Staubli VAL3: io.pjx

--- io.pjx ---
Parameters version=s8.10.3Cs9_BS2093 stackSize=5000 millimeterUnit=true
Program file=commentIO.pgx
Program file=getAnaIO.pgx
Program file=getAngIOSize.pgx
Program file=getDigIO.pgx
Program file=getDigIOSize.pgx
Program file=init.pgx
Program file=linkIO.pgx
Program file=linkStatusIO.pgx
Program file=resetBusSelect.pgx
Program file=setAnaOutput.pgx
Program file=setAngINList.pgx
Program file=setAngOUTList.pgx
Program file=setDigOutNoAlm.pgx
Program file=setDigOutput.pgx
Program file=start.pgx
Program file=stop.pgx
Program file=waitAnaInput.pgx
Program file=waitDigInput.pgx
Data file=io.dtx
Library alias=rs path=Disk://source/projectSource/robotStatus/robotStatus.pjx
Type name=dioItem path=Disk://source/template/dioItem/dioItem.pjx
Type name=aioItem path=Disk://source/template/aioItem/aioItem.pjx

--- io.dtx ---
public aio _aInEthercat[16]
public aio _aInEthernet[20]
public aio _aInModbus[16]
public aio _aInProfibus[16]
public aio _aInProfinet[8]
  [0] = {link=61F414E4-CB2A-4A4A-A70F-3C6D612AB3AA}
  [1] = {link=443D484E-60E0-45BD-99C4-97873755DFDA}
  [2] = {link=73C25A3F-C0C4-4812-B693-CDA309C2D933}
  [3] = {link=D3F549A9-B3EA-403D-BF4C-7070E9F5D37B}
  [4] = {link=F3F4C9C0-1F7C-4DDD-AA59-2014D98A0E36}
  [5] = {link=64B8C6E8-3A71-49B0-BD71-5728B0329AAB}
  [6] = {link=218C656F-9E2A-4E1B-B485-E83EC4F0FE99}
  [7] = {link=66AABE0A-89B4-481F-83AB-C514130625BA}
public aio _aInUser[16]
public aio _aOEthercat[16]
public aio _aOEthernet[20]
public aio _aOModbus[16]
public aio _aOProfibus[16]
public aio _aOProfinet[8]
  [0] = {link=5FFE21EC-528D-4C47-A8D5-7C4CFC474629}
  [1] = {link=6C0C10F5-5D52-4306-AECC-A9DCF4E15FA5}
  [2] = {link=96FBB4C4-7B28-4C73-AFB9-CDBD1E0FA505}
  [3] = {link=3CD60215-4462-490B-9BA1-05C4B27AD9CF}
  [4] = {link=45C44C09-08B8-4891-969D-45390D63770F}
  [5] = {link=DD02F8D1-5F5E-4FDF-BD15-7DB79F0068FE}
  [6] = {link=0578226E-4341-48AC-B576-D095F8D3C1C5}
  [7] = {link=D8473422-71DA-4369-901E-04429E7E73E1}
public aio _aOutUser[16]
public aio aInJobNumber
public aio aInVirtual[24]
  [0] = {link=VirtualIOBoards\VirtualBoard0\%IF128}
  [1] = {link=VirtualIOBoards\VirtualBoard0\%IF160}
  [2] = {link=VirtualIOBoards\VirtualBoard0\%IF192}
  [3] = {link=VirtualIOBoards\VirtualBoard0\%IF224}
  [4] = {link=VirtualIOBoards\VirtualBoard0\%IF256}
  [5] = {link=VirtualIOBoards\VirtualBoard0\%IF288}
  [6] = {link=VirtualIOBoards\VirtualBoard0\%IF320}
  [7] = {link=VirtualIOBoards\VirtualBoard0\%IF352}
  [8] = {link=VirtualIOBoards\VirtualBoard0\%IF384}
  [9] = {link=VirtualIOBoards\VirtualBoard0\%IF416}
  [10] = {link=VirtualIOBoards\VirtualBoard0\%IF448}
  [11] = {link=VirtualIOBoards\VirtualBoard0\%IF480}
  [12] = {link=VirtualIOBoards\VirtualBoard0\%IF512}
  [13] = {link=VirtualIOBoards\VirtualBoard0\%IF544}
  [14] = {link=VirtualIOBoards\VirtualBoard0\%IF576}
  [15] = {link=VirtualIOBoards\VirtualBoard0\%IF608}
  [16] = {link=VirtualIOBoards\VirtualBoard0\%IF640}
  [17] = {link=VirtualIOBoards\VirtualBoard0\%IF672}
  [18] = {link=VirtualIOBoards\VirtualBoard0\%IF704}
  [19] = {link=VirtualIOBoards\VirtualBoard0\%IF736}
  [20] = {link=VirtualIOBoards\VirtualBoard0\%IF768}
  [21] = {link=VirtualIOBoards\VirtualBoard0\%IF800}
  [22] = {link=VirtualIOBoards\VirtualBoard0\%IF832}
  [23] = {link=VirtualIOBoards\VirtualBoard0\%IF864}
public aio aInput[8]
  [0] = {link=61F414E4-CB2A-4A4A-A70F-3C6D612AB3AA}
  [1] = {link=443D484E-60E0-45BD-99C4-97873755DFDA}
  [2] = {link=73C25A3F-C0C4-4812-B693-CDA309C2D933}
  [3] = {link=D3F549A9-B3EA-403D-BF4C-7070E9F5D37B}
  [4] = {link=F3F4C9C0-1F7C-4DDD-AA59-2014D98A0E36}
  [5] = {link=64B8C6E8-3A71-49B0-BD71-5728B0329AAB}
  [6] = {link=218C656F-9E2A-4E1B-B485-E83EC4F0FE99}
  [7] = {link=66AABE0A-89B4-481F-83AB-C514130625BA}
public aio aOutJobNumber
public aio aOutVirtual[24]
  [0] = {link=VirtualIOBoards\VirtualBoard0\%QF128}
  [1] = {link=VirtualIOBoards\VirtualBoard0\%QF160}
  [2] = {link=VirtualIOBoards\VirtualBoard0\%QF192}
  [3] = {link=VirtualIOBoards\VirtualBoard0\%QF224}
  [4] = {link=VirtualIOBoards\VirtualBoard0\%QF256}
  [5] = {link=VirtualIOBoards\VirtualBoard0\%QF288}
  [6] = {link=VirtualIOBoards\VirtualBoard0\%QF320}
  [7] = {link=VirtualIOBoards\VirtualBoard0\%QF352}
  [8] = {link=VirtualIOBoards\VirtualBoard0\%QF384}
  [9] = {link=VirtualIOBoards\VirtualBoard0\%QF416}
  [10] = {link=VirtualIOBoards\VirtualBoard0\%QF448}
  [11] = {link=VirtualIOBoards\VirtualBoard0\%QF480}
  [12] = {link=VirtualIOBoards\VirtualBoard0\%QF512}
  [13] = {link=VirtualIOBoards\VirtualBoard0\%QF544}
  [14] = {link=VirtualIOBoards\VirtualBoard0\%QF576}
  [15] = {link=VirtualIOBoards\VirtualBoard0\%QF608}
  [16] = {link=VirtualIOBoards\VirtualBoard0\%QF640}
  [17] = {link=VirtualIOBoards\VirtualBoard0\%QF672}
  [18] = {link=VirtualIOBoards\VirtualBoard0\%QF704}
  [19] = {link=VirtualIOBoards\VirtualBoard0\%QF736}
  [20] = {link=VirtualIOBoards\VirtualBoard0\%QF768}
  [21] = {link=VirtualIOBoards\VirtualBoard0\%QF800}
  [22] = {link=VirtualIOBoards\VirtualBoard0\%QF832}
  [23] = {link=VirtualIOBoards\VirtualBoard0\%QF864}
public aio aOutput[8]
  [0] = {link=5FFE21EC-528D-4C47-A8D5-7C4CFC474629}
  [1] = {link=6C0C10F5-5D52-4306-AECC-A9DCF4E15FA5}
  [2] = {link=96FBB4C4-7B28-4C73-AFB9-CDBD1E0FA505}
  [3] = {link=3CD60215-4462-490B-9BA1-05C4B27AD9CF}
  [4] = {link=45C44C09-08B8-4891-969D-45390D63770F}
  [5] = {link=DD02F8D1-5F5E-4FDF-BD15-7DB79F0068FE}
  [6] = {link=0578226E-4341-48AC-B576-D095F8D3C1C5}
  [7] = {link=D8473422-71DA-4369-901E-04429E7E73E1}
public aioItem aInItem[8]
  [0]
    aio aAio = {link=61F414E4-CB2A-4A4A-A70F-3C6D612AB3AA}
    string sComment = "接收程序号"
  [1]
    aio aAio = {link=443D484E-60E0-45BD-99C4-97873755DFDA}
    string sComment = "刷子号反馈"
  [2]
    aio aAio = {link=73C25A3F-C0C4-4812-B693-CDA309C2D933}
    string sComment = "备用"
  [3]
    aio aAio = {link=D3F549A9-B3EA-403D-BF4C-7070E9F5D37B}
    string sComment = "备用"
  [4]
    aio aAio = {link=F3F4C9C0-1F7C-4DDD-AA59-2014D98A0E36}
    string sComment = "备用"
  [5]
    aio aAio = {link=64B8C6E8-3A71-49B0-BD71-5728B0329AAB}
    string sComment = "备用"
  [6]
    aio aAio = {link=218C656F-9E2A-4E1B-B485-E83EC4F0FE99}
    string sComment = "备用"
  [7]
    aio aAio = {link=66AABE0A-89B4-481F-83AB-C514130625BA}
    string sComment = "备用"
public aioItem aOutItem[8]
  [0]
    aio aAio = {link=5FFE21EC-528D-4C47-A8D5-7C4CFC474629}
    string sComment = "程序号反馈"
  [1]
    aio aAio = {link=6C0C10F5-5D52-4306-AECC-A9DCF4E15FA5}
    string sComment = "刷子号"
  [2]
    aio aAio = {link=96FBB4C4-7B28-4C73-AFB9-CDBD1E0FA505}
    string sComment = "备用"
  [3]
    aio aAio = {link=3CD60215-4462-490B-9BA1-05C4B27AD9CF}
    string sComment = "备用"
  [4]
    aio aAio = {link=45C44C09-08B8-4891-969D-45390D63770F}
    string sComment = "备用"
  [5]
    aio aAio = {link=DD02F8D1-5F5E-4FDF-BD15-7DB79F0068FE}
    string sComment = "备用"
  [6]
    aio aAio = {link=0578226E-4341-48AC-B576-D095F8D3C1C5}
    string sComment = "备用"
  [7]
    aio aAio = {link=D8473422-71DA-4369-901E-04429E7E73E1}
    string sComment = "备用"
bool bBusSelect[6]
bool bUseAnalog = true
public dio _dInEtherCat[96]
public dio _dInEtherNet[128]
  [0] = {link=3C99ACBA-F1D4-4A68-A21C-89A8C66262F3}
  [1] = {link=A8C10724-75A9-4217-88F5-3321E2E2ACAD}
  [2] = {link=3FECD266-02DB-40D3-AA00-852A922114D7}
  [3] = {link=527ABC03-504A-4B4E-8384-0B648B30A7EE}
  [4] = {link=F6BC421B-A283-4F49-B66E-4A61065D35DB}
  [5] = {link=AF78B140-D810-4E0E-A464-37CD3BF21C1F}
  [6] = {link=54025B48-0E34-4C00-83F4-7C1C00C78D0E}
  [7] = {link=C893EABF-80A0-4CC4-8CB1-35D77AC88EDF}
  [8] = {link=B91BA001-E4EA-48BD-931D-F38D504579C9}
  [9] = {link=F2BD5778-F2D0-400E-8EB0-EB74F7A1D168}
  [10] = {link=00F50513-209B-4FEC-BCA0-2732338E58E1}
  [11] = {link=881EE622-97CE-4B32-A64C-C6F69EF3ED05}
  [12] = {link=56AD774C-0018-466F-B601-292CE44541BC}
  [13] = {link=4324DB33-706B-4D11-8D24-EAF877265392}
  [14] = {link=5AF359B1-8E78-40AA-A03B-F8A0077C8703}
  [15] = {link=ApplicomIO-1\PFN-IN\%I0[15]}
  [16] = {link=ApplicomIO-1\PFN-IN\%I0[16]}
  [17] = {link=ApplicomIO-1\PFN-IN\%I0[17]}
  [18] = {link=ApplicomIO-1\PFN-IN\%I0[18]}
  [19] = {link=ApplicomIO-1\PFN-IN\%I0[19]}
  [20] = {link=ApplicomIO-1\PFN-IN\%I0[20]}
  [21] = {link=ApplicomIO-1\PFN-IN\%I0[21]}
  [22] = {link=ApplicomIO-1\PFN-IN\%I0[22]}
  [23] = {link=ApplicomIO-1\PFN-IN\%I0[23]}
  [24] = {link=ApplicomIO-1\PFN-IN\%I0[24]}
  [25] = {link=ApplicomIO-1\PFN-IN\%I0[25]}
  [26] = {link=ApplicomIO-1\PFN-IN\%I0[26]}
  [27] = {link=ApplicomIO-1\PFN-IN\%I0[27]}
  [28] = {link=ApplicomIO-1\PFN-IN\%I0[28]}
  [29] = {link=ApplicomIO-1\PFN-IN\%I0[29]}
  [30] = {link=ApplicomIO-1\PFN-IN\%I0[30]}
  [31] = {link=ApplicomIO-1\PFN-IN\%I0[31]}
  [32] = {link=ApplicomIO-1\PFN-IN\%I0[32]}
  [33] = {link=ApplicomIO-1\PFN-IN\%I0[33]}
  [34] = {link=ApplicomIO-1\PFN-IN\%I0[34]}
  [35] = {link=ApplicomIO-1\PFN-IN\%I0[35]}
  [36] = {link=ApplicomIO-1\PFN-IN\%I0[36]}
  [37] = {link=ApplicomIO-1\PFN-IN\%I0[37]}
  [38] = {link=ApplicomIO-1\PFN-IN\%I0[38]}
  [39] = {link=ApplicomIO-1\PFN-IN\%I0[39]}
  [40] = {link=ApplicomIO-1\PFN-IN\%I0[40]}
  [41] = {link=ApplicomIO-1\PFN-IN\%I0[41]}
  [42] = {link=ApplicomIO-1\PFN-IN\%I0[42]}
  [43] = {link=ApplicomIO-1\PFN-IN\%I0[43]}
  [44] = {link=ApplicomIO-1\PFN-IN\%I0[44]}
  [45] = {link=ApplicomIO-1\PFN-IN\%I0[45]}
  [46] = {link=ApplicomIO-1\PFN-IN\%I0[46]}
  [47] = {link=ApplicomIO-1\PFN-IN\%I0[47]}
  [48] = {link=ApplicomIO-1\PFN-IN\%I0[48]}
  [49] = {link=ApplicomIO-1\PFN-IN\%I0[49]}
  [50] = {link=ApplicomIO-1\PFN-IN\%I0[50]}
  [51] = {link=ApplicomIO-1\PFN-IN\%I0[51]}
  [52] = {link=ApplicomIO-1\PFN-IN\%I0[52]}
  [53] = {link=ApplicomIO-1\PFN-IN\%I0[53]}
  [54] = {link=ApplicomIO-1\PFN-IN\%I0[54]}
  [55] = {link=ApplicomIO-1\PFN-IN\%I0[55]}
  [56] = {link=ApplicomIO-1\PFN-IN\%I0[56]}
  [57] = {link=ApplicomIO-1\PFN-IN\%I0[57]}
  [58] = {link=ApplicomIO-1\PFN-IN\%I0[58]}
  [59] = {link=ApplicomIO-1\PFN-IN\%I0[59]}
  [60] = {link=ApplicomIO-1\PFN-IN\%I0[60]}
  [61] = {link=ApplicomIO-1\PFN-IN\%I0[61]}
  [62] = {link=ApplicomIO-1\PFN-IN\%I0[62]}
  [63] = {link=ApplicomIO-1\PFN-IN\%I0[63]}
public dio _dInModbus[96]
public dio _dInProfibus[96]
  [0] = {link=ApplicomIO-1\PFB-BLOCK\%I0[0]}
  [1] = {link=ApplicomIO-1\PFB-BLOCK\%I0[1]}
  [2] = {link=ApplicomIO-1\PFB-BLOCK\%I0[2]}
  [3] = {link=ApplicomIO-1\PFB-BLOCK\%I0[3]}
  [4] = {link=ApplicomIO-1\PFB-BLOCK\%I0[4]}
  [5] = {link=ApplicomIO-1\PFB-BLOCK\%I0[5]}
  [6] = {link=ApplicomIO-1\PFB-BLOCK\%I0[6]}
  [7] = {link=ApplicomIO-1\PFB-BLOCK\%I0[7]}
  [8] = {link=ApplicomIO-1\PFB-BLOCK\%I0[8]}
  [9] = {link=ApplicomIO-1\PFB-BLOCK\%I0[9]}
  [10] = {link=ApplicomIO-1\PFB-BLOCK\%I0[10]}
  [11] = {link=ApplicomIO-1\PFB-BLOCK\%I0[11]}
  [12] = {link=ApplicomIO-1\PFB-BLOCK\%I0[12]}
  [13] = {link=ApplicomIO-1\PFB-BLOCK\%I0[13]}
  [14] = {link=ApplicomIO-1\PFB-BLOCK\%I0[14]}
  [15] = {link=ApplicomIO-1\PFB-BLOCK\%I0[15]}
  [16] = {link=ApplicomIO-1\PFB-BLOCK\%I0[16]}
  [17] = {link=ApplicomIO-1\PFB-BLOCK\%I0[17]}
  [18] = {link=ApplicomIO-1\PFB-BLOCK\%I0[18]}
  [19] = {link=ApplicomIO-1\PFB-BLOCK\%I0[19]}
  [20] = {link=ApplicomIO-1\PFB-BLOCK\%I0[20]}
  [21] = {link=ApplicomIO-1\PFB-BLOCK\%I0[21]}
  [22] = {link=ApplicomIO-1\PFB-BLOCK\%I0[22]}
  [23] = {link=ApplicomIO-1\PFB-BLOCK\%I0[23]}
  [24] = {link=ApplicomIO-1\PFB-BLOCK\%I0[24]}
  [25] = {link=ApplicomIO-1\PFB-BLOCK\%I0[25]}
  [26] = {link=ApplicomIO-1\PFB-BLOCK\%I0[26]}
  [27] = {link=ApplicomIO-1\PFB-BLOCK\%I0[27]}
  [28] = {link=ApplicomIO-1\PFB-BLOCK\%I0[28]}
  [29] = {link=ApplicomIO-1\PFB-BLOCK\%I0[29]}
  [30] = {link=ApplicomIO-1\PFB-BLOCK\%I0[30]}
  [31] = {link=ApplicomIO-1\PFB-BLOCK\%I0[31]}
  [32] = {link=ApplicomIO-1\PFB-BLOCK\%I0[32]}
  [33] = {link=ApplicomIO-1\PFB-BLOCK\%I0[33]}
  [34] = {link=ApplicomIO-1\PFB-BLOCK\%I0[34]}
  [35] = {link=ApplicomIO-1\PFB-BLOCK\%I0[35]}
  [36] = {link=ApplicomIO-1\PFB-BLOCK\%I0[36]}
  [37] = {link=ApplicomIO-1\PFB-BLOCK\%I0[37]}
  [38] = {link=ApplicomIO-1\PFB-BLOCK\%I0[38]}
  [39] = {link=ApplicomIO-1\PFB-BLOCK\%I0[39]}
  [40] = {link=ApplicomIO-1\PFB-BLOCK\%I0[40]}
  [41] = {link=ApplicomIO-1\PFB-BLOCK\%I0[41]}
  [42] = {link=ApplicomIO-1\PFB-BLOCK\%I0[42]}
  [43] = {link=ApplicomIO-1\PFB-BLOCK\%I0[43]}
  [44] = {link=ApplicomIO-1\PFB-BLOCK\%I0[44]}
  [45] = {link=ApplicomIO-1\PFB-BLOCK\%I0[45]}
  [46] = {link=ApplicomIO-1\PFB-BLOCK\%I0[46]}
  [47] = {link=ApplicomIO-1\PFB-BLOCK\%I0[47]}
  [48] = {link=ApplicomIO-1\PFB-BLOCK\%I0[48]}
  [49] = {link=ApplicomIO-1\PFB-BLOCK\%I0[49]}
  [50] = {link=ApplicomIO-1\PFB-BLOCK\%I0[50]}
  [51] = {link=ApplicomIO-1\PFB-BLOCK\%I0[51]}
  [52] = {link=ApplicomIO-1\PFB-BLOCK\%I0[52]}
  [53] = {link=ApplicomIO-1\PFB-BLOCK\%I0[53]}
  [54] = {link=ApplicomIO-1\PFB-BLOCK\%I0[54]}
  [55] = {link=ApplicomIO-1\PFB-BLOCK\%I0[55]}
  [56] = {link=ApplicomIO-1\PFB-BLOCK\%I0[56]}
  [57] = {link=ApplicomIO-1\PFB-BLOCK\%I0[57]}
  [58] = {link=ApplicomIO-1\PFB-BLOCK\%I0[58]}
  [59] = {link=ApplicomIO-1\PFB-BLOCK\%I0[59]}
  [60] = {link=ApplicomIO-1\PFB-BLOCK\%I0[60]}
  [61] = {link=ApplicomIO-1\PFB-BLOCK\%I0[61]}
  [62] = {link=ApplicomIO-1\PFB-BLOCK\%I0[62]}
  [63] = {link=ApplicomIO-1\PFB-BLOCK\%I0[63]}
public dio _dInProfinet[128]
  [0] = {link=801699AD-0D4E-40AF-A7AF-E7C40311637E}
  [1] = {link=842E3CE8-5982-430F-AA8E-B2F701DC178B}
  [2] = {link=F299EF97-EDDD-4BB8-AA07-719E60051D06}
  [3] = {link=0D6C59A5-572E-4845-9D24-D0618D782DD4}
  [4] = {link=CC171C2B-47CE-4C45-9659-7FCDC013CE94}
  [5] = {link=1A1317E2-9651-45BA-ACEA-D1820BFA9703}
  [6] = {link=1B720B0E-A94A-4B35-8241-512C8CFE7420}
  [7] = {link=6F68113A-0DD2-4F74-B0DE-02F63C641B3D}
  [8] = {link=DB25555B-9639-404C-BF41-A1E4182E7853}
  [9] = {link=A68ADCD7-077C-45ED-AE36-CA1771248567}
  [10] = {link=3971923C-046E-4FB8-8CDF-8298982DD00B}
  [11] = {link=C253DB67-AB15-493D-BA5F-F7404DA89E40}
  [12] = {link=5F58F424-9E7E-46E6-B5AD-37E850D30CCF}
  [13] = {link=0B266260-B4AD-4902-9CA8-DAC05E19210B}
  [14] = {link=20B44CE4-2E83-403B-A39C-4F8E5CA01265}
  [15] = {link=CD23C02B-CC02-4E28-82D0-6EB1534712A8}
  [16] = {link=550C0093-735F-4929-AB88-92E210EEA585}
  [17] = {link=58675BC9-A902-44A6-9D1E-CDCDD371E5BF}
  [18] = {link=C6C06F3F-E54C-4EE8-B5A1-0B392CB95D19}
  [19] = {link=E7996F97-FFB6-4A1D-8389-FC391F807530}
  [20] = {link=545E5659-957E-409A-983D-845A312BF10F}
  [21] = {link=896C2D61-98DD-43B3-A9FF-B63B82E13F66}
  [22] = {link=CB058ED0-A460-493F-ACD8-83515F19CB22}
  [23] = {link=8EC8BEC8-3882-4E09-82EB-ED6F4043F345}
  [24] = {link=6614FE1F-5D84-418F-8C43-3AD6E08D9885}
  [25] = {link=A0D729AE-192B-4443-98B3-A6978F97C45B}
  [26] = {link=8274EAD0-4711-40CE-9532-B3E4F6D5E848}
  [27] = {link=A4D7A453-0050-4322-BCBB-255C4251B0BA}
  [28] = {link=0CFB91EB-8B07-41BC-89A1-F8BBECCF0624}
  [29] = {link=4F7299CD-79A3-4FE2-8435-19083E83C2B9}
  [30] = {link=E49B7D09-65F8-4955-B810-3C508C434830}
  [31] = {link=2BAB1321-D2BB-48C2-8DEA-1230FF1A9D85}
  [32] = {link=C00D5C02-BF78-4EF5-B868-C5B31E42BE7F}
  [33] = {link=96859C69-E3EF-4F26-913D-E25096C13C5F}
  [34] = {link=7920EEE9-3DBF-43F3-9541-7FBE207ECE53}
  [35] = {link=1DB9160A-F63F-4C13-93B5-492FEDD177E2}
  [36] = {link=1FC4D9B1-EE44-4A9B-A22D-5889BB08EE1E}
  [37] = {link=BF970AFE-565C-4857-97A6-5A54DDAE79B6}
  [38] = {link=F909C748-B7A8-4470-A6FD-BA1A46FE4E68}
  [39] = {link=8517CD21-2BAD-4F53-9136-89235F4060C6}
  [40] = {link=6DDBB7AB-AC7B-4F3D-A091-1238925E0448}
  [41] = {link=C3CF7374-59EF-4029-99B4-FC98E25808BB}
  [42] = {link=90C02E77-8235-444D-99EB-D816EF90AFE5}
  [43] = {link=E44556E2-741A-40A0-89B2-8E32677B3EB1}
  [44] = {link=D8AFCC23-6F61-4ADD-8DE3-3FE1547AD28D}
  [45] = {link=98BC2888-38BC-4A33-A762-BDEC3E36173F}
  [46] = {link=A24DA26D-2F10-46AE-809B-0B04336865AA}
  [47] = {link=04D21FA2-EBE1-4E66-8338-7CB17174A724}
  [48] = {link=E766472B-9569-4911-A858-6F7708718D01}
  [49] = {link=92C360C1-157E-40E1-9184-03D53ECDF3F7}
  [50] = {link=6E33B145-BAC8-48E7-A184-E5A9D90B515B}
  [51] = {link=D5FDB290-CB76-4852-8AF4-F9B6FA5D3E2D}
  [52] = {link=547C3630-B2EA-42F8-AB37-EEB4C81AA149}
  [53] = {link=A60C469C-4F75-4C30-9347-66365041DE79}
  [54] = {link=6E14BCEF-8B69-4038-B259-0EF712D2AB66}
  [55] = {link=B19F0E1B-CE25-49C3-9ED7-92404708DBC9}
  [56] = {link=AFC49D6D-7F53-41F5-8159-6058E9291542}
  [57] = {link=BB08126F-937C-4C50-9A1C-252CB13BB25C}
  [58] = {link=15BF4171-EFAA-47B7-BEF9-A698BE11011C}
  [59] = {link=9A261803-1F52-41D2-8355-1C79BF1BB94D}
  [60] = {link=18F63136-91BD-4FEE-8DA3-2AA9D2E8FFA8}
  [61] = {link=55E89D2C-C808-4026-99D2-85E324C475F9}
  [62] = {link=45535323-0512-46DB-8EB0-4BF3F55D73C7}
  [63] = {link=23943399-CEE5-49D9-BFD9-55B5920F548B}
  [64] = {link=364F41EB-6BA1-4700-BD0A-C2236839044E}
  [65] = {link=96EFCAAE-6B9A-4070-B9EC-2035BA94CCB3}
  [66] = {link=FD79DB68-803F-47E7-8305-8CFFFE519C88}
  [67] = {link=82CF98E3-5511-4523-9501-B4BBAD9DC96D}
  [68] = {link=43A446B7-3C25-4DD5-9597-27365DBE2539}
  [69] = {link=01367322-9745-4163-BFB8-DF881D521F4A}
  [70] = {link=1F635259-38C5-4AB2-B093-ADA4F82FD92B}
  [71] = {link=80065B3A-E7EF-4B6D-A30A-AC2F8A1FF9BD}
  [72] = {link=138692BF-FCCE-4B34-B0E8-8C4B22C67F12}
  [73] = {link=2F598E66-6704-43A6-A433-14D902C15D10}
  [74] = {link=3D7C9642-411B-40D3-B3B9-C83D24259AF4}
  [75] = {link=2E14C0AE-1F04-4256-8959-DEAD28BB69AE}
  [76] = {link=D90512A1-D0E1-41B2-8294-59D7C1ADD8E0}
  [77] = {link=F9EFA2A2-C655-4B55-8F3F-AAE77A6FD751}
  [78] = {link=8C43F822-1313-4C63-84D2-76D62B96A58F}
  [79] = {link=0BE51982-5E8E-4776-A637-0836608FA4D4}
  [80] = {link=5CC26A0C-A759-4F9D-9C90-7643106A4280}
  [81] = {link=6B2348DB-D0C3-44B1-96EA-09FBC0D6D1F3}
  [82] = {link=091DC27E-E2EB-463E-8E4B-08B48E663650}
  [83] = {link=EC5520D5-F711-48B3-AE90-97344DDBEE5C}
  [84] = {link=E02811C8-C36E-4E92-B28C-81A727813C5B}
  [85] = {link=39EB69C5-9612-415D-9A77-D013E3B8CFD4}
  [86] = {link=FD4FFC3C-593A-4304-8BB2-18534DB95237}
  [87] = {link=D2ECCFF1-C6D1-48A4-B3A9-F333711A9798}
  [88] = {link=13EA7043-3380-41E5-9177-AAC787C21C39}
  [89] = {link=5475660F-31B7-47C3-808C-FBAB066EFE6D}
  [90] = {link=93D7CC16-1244-4B9F-85C2-564B516A38A6}
  [91] = {link=A2A5B44E-CAC8-47F1-A810-875EED5095FB}
  [92] = {link=2F9951E4-3414-412E-A45B-55B5D632DA1B}
  [93] = {link=916866A1-8E9C-42B7-A695-7CB9D795E148}
  [94] = {link=CA3200CB-BA9D-4435-B593-6CDDBB86F10C}
  [95] = {link=49AC3AF5-F49B-42A1-90B2-5DB7D6C7E051}
  [96] = {link=64E7B72A-8AE1-43E7-9A21-FF4DABD03910}
  [97] = {link=7BA0757A-43B7-4994-86FC-1740DE8C159E}
  [98] = {link=5ACF5B88-9BD6-435A-8F3F-752FE88E7935}
  [99] = {link=70DFB9C6-9CA4-44C9-8464-A31BA0D039F5}
  [100] = {link=55D5D0F9-E23A-40DA-9955-6BCB63B37099}
  [101] = {link=1AB52030-AE2C-417B-9C38-1633EF57A0DB}
  [102] = {link=FFE2E20E-ABB5-4A36-BE3B-E714CB40E85A}
  [103] = {link=83BC89DD-B780-47A7-BBF0-017BDC2BA365}
  [104] = {link=10D6F5C6-79FE-4371-9CC9-A814346F77C1}
  [105] = {link=240957B0-B56A-4DFB-9281-23480961F3F1}
  [106] = {link=92C2EE73-BB65-4A97-8029-77FB60FFC23C}
  [107] = {link=62C2F98E-E7EB-49ED-971A-83A5444F6152}
  [108] = {link=58CC62E1-4595-401C-8E2F-3122D818CC74}
  [109] = {link=6D2EBC96-6FF5-40C1-83D6-CC8DD3D9FC3A}
  [110] = {link=AEC5DD07-0ABE-4FC2-A89A-ED52FEBBCAD7}
  [111] = {link=D289FF49-1CD8-4174-B7A5-8E375EB48B35}
  [112] = {link=4D3459D2-B2AE-4602-8654-6AD44AA154CE}
  [113] = {link=BE4318FA-0CA3-4B50-ACFD-D0BD90E002BB}
  [114] = {link=03734564-3942-45B2-807F-C861E4A00B4D}
  [115] = {link=18C4B14F-9C0F-4159-B56F-314AFF4BFABC}
  [116] = {link=A703F976-FEB8-4965-8F5A-CAD8585E54F7}
  [117] = {link=F3814F6C-1F81-45E4-8DE4-AB9F0C1AC9C1}
  [118] = {link=CD215C83-5C8C-4339-BF6C-DDE6EDBF5021}
  [119] = {link=295A35FF-B8CC-4A25-BC99-5CC4EFE79E3D}
  [120] = {link=7D822E1A-7C34-46E1-A06C-E10F3FD6B4DE}
  [121] = {link=4A23737B-5C9C-4372-A68A-8F60451AD439}
  [122] = {link=B2909A16-C926-42A5-8387-168FB9DA6D2A}
  [123] = {link=36FA5061-3D34-4793-BCBA-E09767B9821D}
  [124] = {link=0AE8B5A8-7356-480B-AAA1-20AFD496F398}
  [125] = {link=DB043A0E-80EF-4F10-9CBC-7A049A7AEFDE}
  [126] = {link=951CF18F-CA29-47EF-A085-39A8D6CD28C1}
  [127] = {link=6FC2F7D5-08CF-47CC-86FA-1AC31B966FFD}
public dio _dInUser[96]
  [32] = {link=FastIO\fIn0}
  [33] = {link=FastIO\fIn1}
public dio _dOEtherCat[96]
  [0] = {link=EtherCAT-1\%Q0}
  [1] = {link=EtherCAT-1\%Q1}
  [2] = {link=EtherCAT-1\%Q2}
  [3] = {link=EtherCAT-1\%Q3}
  [4] = {link=EtherCAT-1\%Q4}
  [5] = {link=EtherCAT-1\%Q5}
  [6] = {link=EtherCAT-1\%Q6}
  [7] = {link=EtherCAT-1\%Q7}
  [8] = {link=EtherCAT-1\%Q8}
  [9] = {link=EtherCAT-1\%Q9}
  [10] = {link=EtherCAT-1\%Q10}
  [11] = {link=EtherCAT-1\%Q11}
  [12] = {link=EtherCAT-1\%Q12}
  [13] = {link=EtherCAT-1\%Q13}
  [14] = {link=EtherCAT-1\%Q14}
  [15] = {link=EtherCAT-1\%Q15}
  [16] = {link=EtherCAT-1\%Q16}
  [17] = {link=EtherCAT-1\%Q17}
  [18] = {link=EtherCAT-1\%Q18}
  [19] = {link=EtherCAT-1\%Q19}
  [20] = {link=EtherCAT-1\%Q20}
  [21] = {link=EtherCAT-1\%Q21}
  [22] = {link=EtherCAT-1\%Q22}
  [23] = {link=EtherCAT-1\%Q23}
  [24] = {link=EtherCAT-1\%Q24}
  [25] = {link=EtherCAT-1\%Q25}
  [26] = {link=EtherCAT-1\%Q26}
  [27] = {link=EtherCAT-1\%Q27}
  [28] = {link=EtherCAT-1\%Q28}
  [29] = {link=EtherCAT-1\%Q29}
  [30] = {link=EtherCAT-1\%Q30}
  [31] = {link=EtherCAT-1\%Q31}
  [32] = {link=EtherCAT-1\%Q32}
  [33] = {link=EtherCAT-1\%Q33}
  [34] = {link=EtherCAT-1\%Q34}
  [35] = {link=EtherCAT-1\%Q35}
  [36] = {link=EtherCAT-1\%Q36}
  [37] = {link=EtherCAT-1\%Q37}
  [38] = {link=EtherCAT-1\%Q38}
  [39] = {link=EtherCAT-1\%Q39}
  [40] = {link=EtherCAT-1\%Q40}
  [41] = {link=EtherCAT-1\%Q41}
  [42] = {link=EtherCAT-1\%Q42}
  [43] = {link=EtherCAT-1\%Q43}
  [44] = {link=EtherCAT-1\%Q44}
  [45] = {link=EtherCAT-1\%Q45}
  [46] = {link=EtherCAT-1\%Q46}
  [47] = {link=EtherCAT-1\%Q47}
  [48] = {link=EtherCAT-1\%Q48}
  [49] = {link=EtherCAT-1\%Q49}
  [50] = {link=EtherCAT-1\%Q50}
  [51] = {link=EtherCAT-1\%Q51}
  [52] = {link=EtherCAT-1\%Q52}
  [53] = {link=EtherCAT-1\%Q53}
  [54] = {link=EtherCAT-1\%Q54}
  [55] = {link=EtherCAT-1\%Q55}
  [56] = {link=EtherCAT-1\%Q56}
  [57] = {link=EtherCAT-1\%Q57}
  [58] = {link=EtherCAT-1\%Q58}
  [59] = {link=EtherCAT-1\%Q59}
  [60] = {link=EtherCAT-1\%Q60}
  [61] = {link=EtherCAT-1\%Q61}
  [62] = {link=EtherCAT-1\%Q62}
  [63] = {link=EtherCAT-1\%Q63}
public dio _dOEtherNet[128]
  [0] = {link=ApplicomIO-1\PFN-OUT\%Q0[0]}
  [1] = {link=ApplicomIO-1\PFN-OUT\%Q0[1]}
  [2] = {link=ApplicomIO-1\PFN-OUT\%Q0[2]}
  [3] = {link=ApplicomIO-1\PFN-OUT\%Q0[3]}
  [4] = {link=ApplicomIO-1\PFN-OUT\%Q0[4]}
  [5] = {link=ApplicomIO-1\PFN-OUT\%Q0[5]}
  [6] = {link=ApplicomIO-1\PFN-OUT\%Q0[6]}
  [7] = {link=ApplicomIO-1\PFN-OUT\%Q0[7]}
  [8] = {link=ApplicomIO-1\PFN-OUT\%Q0[8]}
  [9] = {link=ApplicomIO-1\PFN-OUT\%Q0[9]}
  [10] = {link=ApplicomIO-1\PFN-OUT\%Q0[10]}
  [11] = {link=ApplicomIO-1\PFN-OUT\%Q0[11]}
  [12] = {link=ApplicomIO-1\PFN-OUT\%Q0[12]}
  [13] = {link=ApplicomIO-1\PFN-OUT\%Q0[13]}
  [14] = {link=ApplicomIO-1\PFN-OUT\%Q0[14]}
  [15] = {link=ApplicomIO-1\PFN-OUT\%Q0[15]}
  [16] = {link=ApplicomIO-1\PFN-OUT\%Q0[16]}
  [17] = {link=ApplicomIO-1\PFN-OUT\%Q0[17]}
  [18] = {link=ApplicomIO-1\PFN-OUT\%Q0[18]}
  [19] = {link=ApplicomIO-1\PFN-OUT\%Q0[19]}
  [20] = {link=ApplicomIO-1\PFN-OUT\%Q0[20]}
  [21] = {link=ApplicomIO-1\PFN-OUT\%Q0[21]}
  [22] = {link=ApplicomIO-1\PFN-OUT\%Q0[22]}
  [23] = {link=ApplicomIO-1\PFN-OUT\%Q0[23]}
  [24] = {link=ApplicomIO-1\PFN-OUT\%Q0[24]}
  [25] = {link=ApplicomIO-1\PFN-OUT\%Q0[25]}
  [26] = {link=ApplicomIO-1\PFN-OUT\%Q0[26]}
  [27] = {link=ApplicomIO-1\PFN-OUT\%Q0[27]}
  [28] = {link=ApplicomIO-1\PFN-OUT\%Q0[28]}
  [29] = {link=ApplicomIO-1\PFN-OUT\%Q0[29]}
  [30] = {link=ApplicomIO-1\PFN-OUT\%Q0[30]}
  [31] = {link=ApplicomIO-1\PFN-OUT\%Q0[31]}
  [32] = {link=ApplicomIO-1\PFN-OUT\%Q0[32]}
  [33] = {link=ApplicomIO-1\PFN-OUT\%Q0[33]}
  [34] = {link=ApplicomIO-1\PFN-OUT\%Q0[34]}
  [35] = {link=ApplicomIO-1\PFN-OUT\%Q0[35]}
  [36] = {link=ApplicomIO-1\PFN-OUT\%Q0[36]}
  [37] = {link=ApplicomIO-1\PFN-OUT\%Q0[37]}
  [38] = {link=ApplicomIO-1\PFN-OUT\%Q0[38]}
  [39] = {link=ApplicomIO-1\PFN-OUT\%Q0[39]}
  [40] = {link=ApplicomIO-1\PFN-OUT\%Q0[40]}
  [41] = {link=ApplicomIO-1\PFN-OUT\%Q0[41]}
  [42] = {link=ApplicomIO-1\PFN-OUT\%Q0[42]}
  [43] = {link=ApplicomIO-1\PFN-OUT\%Q0[43]}
  [44] = {link=ApplicomIO-1\PFN-OUT\%Q0[44]}
  [45] = {link=ApplicomIO-1\PFN-OUT\%Q0[45]}
  [46] = {link=ApplicomIO-1\PFN-OUT\%Q0[46]}
  [47] = {link=ApplicomIO-1\PFN-OUT\%Q0[47]}
  [48] = {link=ApplicomIO-1\PFN-OUT\%Q0[48]}
  [49] = {link=ApplicomIO-1\PFN-OUT\%Q0[49]}
  [50] = {link=ApplicomIO-1\PFN-OUT\%Q0[50]}
  [51] = {link=ApplicomIO-1\PFN-OUT\%Q0[51]}
  [52] = {link=ApplicomIO-1\PFN-OUT\%Q0[52]}
  [53] = {link=ApplicomIO-1\PFN-OUT\%Q0[53]}
  [54] = {link=ApplicomIO-1\PFN-OUT\%Q0[54]}
  [55] = {link=ApplicomIO-1\PFN-OUT\%Q0[55]}
  [56] = {link=ApplicomIO-1\PFN-OUT\%Q0[56]}
  [57] = {link=ApplicomIO-1\PFN-OUT\%Q0[57]}
  [58] = {link=ApplicomIO-1\PFN-OUT\%Q0[58]}
  [59] = {link=ApplicomIO-1\PFN-OUT\%Q0[59]}
  [60] = {link=ApplicomIO-1\PFN-OUT\%Q0[60]}
  [61] = {link=ApplicomIO-1\PFN-OUT\%Q0[61]}
  [62] = {link=ApplicomIO-1\PFN-OUT\%Q0[62]}
  [63] = {link=ApplicomIO-1\PFN-OUT\%Q0[63]}
public dio _dOModbus[96]
public dio _dOProfibus[96]
  [0] = {link=ApplicomIO-1\PFB-BLOCK\%Q0[0]}
  [1] = {link=ApplicomIO-1\PFB-BLOCK\%Q0[1]}
  [2] = {link=ApplicomIO-1\PFB-BLOCK\%Q0[2]}
  [3] = {link=ApplicomIO-1\PFB-BLOCK\%Q0[3]}
  [4] = {link=ApplicomIO-1\PFB-BLOCK\%Q0[4]}
  [5] = {link=ApplicomIO-1\PFB-BLOCK\%Q0[5]}
  [6] = {link=ApplicomIO-1\PFB-BLOCK\%Q0[6]}
  [7] = {link=ApplicomIO-1\PFB-BLOCK\%Q0[7]}
  [8] = {link=ApplicomIO-1\PFB-BLOCK\%Q0[8]}
  [9] = {link=ApplicomIO-1\PFB-BLOCK\%Q0[9]}
  [10] = {link=ApplicomIO-1\PFB-BLOCK\%Q0[10]}
  [11] = {link=ApplicomIO-1\PFB-BLOCK\%Q0[11]}
  [12] = {link=ApplicomIO-1\PFB-BLOCK\%Q0[12]}
  [13] = {link=ApplicomIO-1\PFB-BLOCK\%Q0[13]}
  [14] = {link=ApplicomIO-1\PFB-BLOCK\%Q0[14]}
  [15] = {link=ApplicomIO-1\PFB-BLOCK\%Q0[15]}
  [16] = {link=ApplicomIO-1\PFB-BLOCK\%Q0[16]}
  [17] = {link=ApplicomIO-1\PFB-BLOCK\%Q0[17]}
  [18] = {link=ApplicomIO-1\PFB-BLOCK\%Q0[18]}
  [19] = {link=ApplicomIO-1\PFB-BLOCK\%Q0[19]}
  [20] = {link=ApplicomIO-1\PFB-BLOCK\%Q0[20]}
  [21] = {link=ApplicomIO-1\PFB-BLOCK\%Q0[21]}
  [22] = {link=ApplicomIO-1\PFB-BLOCK\%Q0[22]}
  [23] = {link=ApplicomIO-1\PFB-BLOCK\%Q0[23]}
  [24] = {link=ApplicomIO-1\PFB-BLOCK\%Q0[24]}
  [25] = {link=ApplicomIO-1\PFB-BLOCK\%Q0[25]}
  [26] = {link=ApplicomIO-1\PFB-BLOCK\%Q0[26]}
  [27] = {link=ApplicomIO-1\PFB-BLOCK\%Q0[27]}
  [28] = {link=ApplicomIO-1\PFB-BLOCK\%Q0[28]}
  [29] = {link=ApplicomIO-1\PFB-BLOCK\%Q0[29]}
  [30] = {link=ApplicomIO-1\PFB-BLOCK\%Q0[30]}
  [31] = {link=ApplicomIO-1\PFB-BLOCK\%Q0[31]}
  [32] = {link=ApplicomIO-1\PFB-BLOCK\%Q0[32]}
  [33] = {link=ApplicomIO-1\PFB-BLOCK\%Q0[33]}
  [34] = {link=ApplicomIO-1\PFB-BLOCK\%Q0[34]}
  [35] = {link=ApplicomIO-1\PFB-BLOCK\%Q0[35]}
  [36] = {link=ApplicomIO-1\PFB-BLOCK\%Q0[36]}
  [37] = {link=ApplicomIO-1\PFB-BLOCK\%Q0[37]}
  [38] = {link=ApplicomIO-1\PFB-BLOCK\%Q0[38]}
  [39] = {link=ApplicomIO-1\PFB-BLOCK\%Q0[39]}
  [40] = {link=ApplicomIO-1\PFB-BLOCK\%Q0[40]}
  [41] = {link=ApplicomIO-1\PFB-BLOCK\%Q0[41]}
  [42] = {link=ApplicomIO-1\PFB-BLOCK\%Q0[42]}
  [43] = {link=ApplicomIO-1\PFB-BLOCK\%Q0[43]}
  [44] = {link=ApplicomIO-1\PFB-BLOCK\%Q0[44]}
  [45] = {link=ApplicomIO-1\PFB-BLOCK\%Q0[45]}
  [46] = {link=ApplicomIO-1\PFB-BLOCK\%Q0[46]}
  [47] = {link=ApplicomIO-1\PFB-BLOCK\%Q0[47]}
  [48] = {link=ApplicomIO-1\PFB-BLOCK\%Q0[48]}
  [49] = {link=ApplicomIO-1\PFB-BLOCK\%Q0[49]}
  [50] = {link=ApplicomIO-1\PFB-BLOCK\%Q0[50]}
  [51] = {link=ApplicomIO-1\PFB-BLOCK\%Q0[51]}
  [52] = {link=ApplicomIO-1\PFB-BLOCK\%Q0[52]}
  [53] = {link=ApplicomIO-1\PFB-BLOCK\%Q0[53]}
  [54] = {link=ApplicomIO-1\PFB-BLOCK\%Q0[54]}
  [55] = {link=ApplicomIO-1\PFB-BLOCK\%Q0[55]}
  [56] = {link=ApplicomIO-1\PFB-BLOCK\%Q0[56]}
  [57] = {link=ApplicomIO-1\PFB-BLOCK\%Q0[57]}
  [58] = {link=ApplicomIO-1\PFB-BLOCK\%Q0[58]}
  [59] = {link=ApplicomIO-1\PFB-BLOCK\%Q0[59]}
  [60] = {link=ApplicomIO-1\PFB-BLOCK\%Q0[60]}
  [61] = {link=ApplicomIO-1\PFB-BLOCK\%Q0[61]}
  [62] = {link=ApplicomIO-1\PFB-BLOCK\%Q0[62]}
  [63] = {link=ApplicomIO-1\PFB-BLOCK\%Q0[63]}
public dio _dOProfinet[128]
  [0] = {link=813E3F4B-A1DE-4C5D-8EAB-0242B6D8A546}
  [1] = {link=364EC08F-C077-495B-A954-158507D3C26C}
  [2] = {link=289A5E8D-11F3-4BEB-8FA4-200735E3A2B7}
  [3] = {link=79705501-C546-4790-A460-3F340ADFDE5C}
  [4] = {link=75D4F3C1-C356-4EDA-B423-02C90835EA7D}
  [5] = {link=3F319035-E82A-4D07-9742-3AFC501B53DF}
  [6] = {link=1CC4B59E-3D71-495F-A34B-473B0A37D044}
  [7] = {link=2087A18A-21B3-4E9A-90F0-0A72D013BBC2}
  [8] = {link=93BF17B5-5C7E-43C6-9C42-3B6025772815}
  [9] = {link=16CB4CF9-3A13-4F09-B6E9-D967DFB15E25}
  [10] = {link=734EBAF3-2CA8-4D3F-A8BB-E168C1322725}
  [11] = {link=07A4EEA8-4CAE-47C3-9487-42EFEC0C0C8E}
  [12] = {link=63159677-63A9-4936-A8C6-E65B2885D59F}
  [13] = {link=698A0489-9B90-43A7-B0CD-777095A36007}
  [14] = {link=C4522756-21A9-4D8A-B398-209F6EFB0977}
  [15] = {link=E3974102-9CCD-497B-BD29-7D9DDF1F0662}
  [16] = {link=D7E9BDA6-AD73-4469-BD4D-C9D8F1711105}
  [17] = {link=C0E9CDD3-3C86-4E8A-BB76-29DD4E724269}
  [18] = {link=19A15CFF-CD59-4687-8101-878C6D297AD0}
  [19] = {link=F886CB4C-7C2D-4AEE-8DA8-19CCB8826A1C}
  [20] = {link=44B2E852-2BDD-46AD-B032-142EDC75806B}
  [21] = {link=E6202C42-8108-4A9C-988A-BA326395584A}
  [22] = {link=4A293BE2-BE94-462E-ACFA-7E01BA496DDB}
  [23] = {link=C4CC4269-4D2F-4B53-89D1-5B6F0F9E20C5}
  [24] = {link=976E4904-0F44-43DA-867D-0C06FC7F067A}
  [25] = {link=26F2F168-65FE-450B-BE6F-27BCBE8A7C37}
  [26] = {link=58979B7C-3302-40C0-9293-D8BDE318359F}
  [27] = {link=32E62FFE-3CE0-449B-8ADB-B460A9E5DE54}
  [28] = {link=1778E8D0-D57F-4F6E-A6A4-A7E0DC8A5FDF}
  [29] = {link=BB6EEE31-C681-41BA-8160-A41199CEAD02}
  [30] = {link=58577585-C0FF-479D-B4D2-FF8F04E87201}
  [31] = {link=E4789C35-874D-4E09-8AF9-741C03AAD9B4}
  [32] = {link=AB4C11BC-0698-4F05-9F77-33C54B19FD7D}
  [33] = {link=A971CAAA-D369-4C08-BB4B-F444CDC4D2F0}
  [34] = {link=EE574E0A-35B5-4DE1-8C9E-C0DF9CDCDFE6}
  [35] = {link=7532402E-1B90-4BA9-83CA-579B1F726874}
  [36] = {link=6F6C7C8F-8851-47C2-9B8E-D33C24B9D39F}
  [37] = {link=4A5CAAE4-C9CD-4421-94AD-56079246CA39}
  [38] = {link=EB7E2C34-F887-4C3F-97E0-01834D630C5E}
  [39] = {link=BDBB409A-6EC7-4423-9FF9-A638D02BF80E}
  [40] = {link=E136414E-B9B9-4DA1-8541-C1A78F1E80BF}
  [41] = {link=8E4798E6-5BA8-40FC-8B4C-D83695D2AB51}
  [42] = {link=28472F68-DF34-4C50-9023-A219CE2C4B1B}
  [43] = {link=1DB5BD39-DE07-40ED-B700-8C7874B04DB0}
  [44] = {link=88484DFD-5685-4FE3-BD11-1467A80C9B34}
  [45] = {link=2F5F1623-83AA-4A31-A803-F6FA4D4BE14A}
  [46] = {link=519B5132-0D61-4FA5-ABD4-96724AED25E8}
  [47] = {link=661BE778-7099-413C-A47D-EC9A4ECEF23E}
  [48] = {link=53B2124C-FE98-440B-9A3D-84530B55B740}
  [49] = {link=229E980F-A7B4-4859-9EE1-BA541F4B5A16}
  [50] = {link=1FA4F26D-23CC-42E9-A819-02B2DD7006DA}
  [51] = {link=2AEDD394-CA8D-4F24-A299-43D2A058ACD5}
  [52] = {link=C28EB1DF-BACA-4254-A598-B532E330438E}
  [53] = {link=E7F3183B-4DF3-459A-ADF7-79D82988755C}
  [54] = {link=2614E536-799A-40AF-9560-80A760021F62}
  [55] = {link=757B7056-4991-459D-8227-2BCDF4BE047B}
  [56] = {link=8C99F1DA-9DA9-4BDF-B60F-FD54ABC54EFA}
  [57] = {link=5AA809C1-68E1-4A24-9F04-C8074121C64A}
  [58] = {link=4A164529-4FC6-4374-9AB6-7CFCFB13974B}
  [59] = {link=70724C45-B1FB-42FE-A3A2-C0AB8AA81684}
  [60] = {link=9EE71F53-97CD-4882-A49E-A6F1E8BC9441}
  [61] = {link=81277848-FDAC-47B2-B4F0-EFE16B2F5C1C}
  [62] = {link=E56352E6-5F75-449C-AD2C-249D38B077FB}
  [63] = {link=5728C013-0742-4355-8E61-1A03F1F076E6}
  [64] = {link=04B33B81-599B-4BDE-99DF-EEC79DF42297}
  [65] = {link=D5C4F9D4-602E-45CC-A360-A9C8DFC51706}
  [66] = {link=0F23F4DE-A6DC-48A8-BD13-38096E17E4BC}
  [67] = {link=725D593E-3E8C-49B9-A0C8-EC5E7EDBEF47}
  [68] = {link=D80F8BA0-A9D7-467A-84F3-2EF911086F28}
  [69] = {link=290333BB-E8D8-473B-B7DA-1770BF97A3BA}
  [70] = {link=3451ABCB-1CE5-49F5-8053-7E43529834C5}
  [71] = {link=1C486D5A-1AEA-494E-AC84-6CEA9FC0F052}
  [72] = {link=0B5202A6-62EE-4D6C-8E76-4A396B266DA1}
  [73] = {link=07376469-6AEC-4E90-A30D-02A336A51CCF}
  [74] = {link=9C60D734-A29B-44DA-837E-97A014720D64}
  [75] = {link=F6F5CEBA-7A13-4322-B86E-E02B17A52B8C}
  [76] = {link=034F848A-A2B4-4107-BA29-37F2DF0B4836}
  [77] = {link=2D3AB11E-A0E7-43D6-A64B-B19DE4EDCA54}
  [78] = {link=6B87E34F-9D7F-4178-ADAD-CF451768FAD1}
  [79] = {link=0BECC0A6-11C6-443C-B8B7-B823C5449F03}
  [80] = {link=0FAFA963-6C61-46BA-8B8E-FD5D821CED0B}
  [81] = {link=E858B3E5-8FFB-4B3B-9E73-58A45F891801}
  [82] = {link=52490A38-A31A-4D56-AA93-4E3292557F7F}
  [83] = {link=07DE5AAD-9C80-4970-8E40-B99AD098B2C3}
  [84] = {link=E76E3858-8352-4107-BC87-39491D8B651A}
  [85] = {link=2B09FA37-BF2E-4ED9-B53F-09BB42630F57}
  [86] = {link=C0D4BCE7-AA67-4991-AD3B-5583CCFF9A80}
  [87] = {link=BBA329F0-9B99-401C-B2C0-5AA54B82A434}
  [88] = {link=1FF771B4-EE27-450D-A9DB-7E394712BF39}
  [89] = {link=19978664-DA67-4FAE-9478-F6C2FD7BC1A1}
  [90] = {link=B280086E-4E78-4C33-A16A-5103EDFD12BA}
  [91] = {link=66D76411-AF4D-465C-BF45-D26D600CE49D}
  [92] = {link=CF5BF486-B482-4F9A-936E-D7550E22D48F}
  [93] = {link=47EF2689-3337-4012-BAD2-52612379B15C}
  [94] = {link=9BC9630D-0782-4292-B056-6CBDA421EF62}
  [95] = {link=CAFB5CCA-B450-480D-9CAD-A29B903F45A9}
  [96] = {link=DCBA4C7F-A728-4F25-89A5-B6259619A80B}
  [97] = {link=6753AC4A-51FA-413E-B4B2-137174F0D507}
  [98] = {link=81370562-9275-47C1-93C0-CB31297CDD20}
  [99] = {link=E6DCC6F0-C964-47CD-B4D7-1BD8BFDA33AE}
  [100] = {link=18C334B4-AE06-448E-96BF-3CD280A2541B}
  [101] = {link=15B48D0D-C668-47AF-A704-10BA0ED6FFE7}
  [102] = {link=DA2930BB-B07C-4C38-ADBB-0FDC55ECF2BB}
  [103] = {link=8DDD8F2E-B5A8-4F54-BD1B-48D04A96C878}
  [104] = {link=72245E17-FF99-4704-8474-EDB79B027BF9}
  [105] = {link=BCF85E34-592F-4BA5-AE76-F1E8F2FD96C1}
  [106] = {link=9ED9CFBB-1644-41A9-955E-D6E7EB6EF2F1}
  [107] = {link=5A6FDD52-29C6-40B7-B97D-88DE84ED4E53}
  [108] = {link=8E4836F5-8A3D-4937-90E9-0F98CBF16A27}
  [109] = {link=4305B788-10E3-4C38-9835-3E94A9820D41}
  [110] = {link=152B6212-6AC5-4D19-A5F9-C32452DCD0BD}
  [111] = {link=60BD22D0-03A0-4632-85E7-7AB9A7B5E9EE}
  [112] = {link=617AC81D-63D2-418A-A221-1A45E82E8F33}
  [113] = {link=DA60158B-5C4B-4C1D-9AEB-3A4C25735862}
  [114] = {link=7E45E59A-6E5F-4DD8-8E87-A62787B5121D}
  [115] = {link=302676B4-AFEF-4A5D-9D0F-7D7EEE15BD09}
  [116] = {link=94FD2E61-B0C4-426E-8CB5-3D13DE4E72D1}
  [117] = {link=5441B2EB-7737-420D-A838-CB6BC6A9AA98}
  [118] = {link=D70A9639-74F8-485B-B1AE-A12B6619BE09}
  [119] = {link=3C4D5DF3-3DD0-4928-9BAC-FF9DB40E9304}
  [120] = {link=389B2383-01D9-4D6D-8093-13CF39736E4D}
  [121] = {link=9C61CF1A-5A0B-480F-A9AF-E365017F4409}
  [122] = {link=D6F4FFC6-5A52-44AE-AAFC-981F5DBD7076}
  [123] = {link=3768B870-3C40-471D-B639-CE39EBCB3865}
  [124] = {link=FCBA4290-2AF9-4EDB-AAB3-C3D5B2BC56ED}
  [125] = {link=FEB8E5C1-4C55-454A-AACA-1D927BE28924}
  [126] = {link=C97B50B1-B825-4E71-A20E-3BFEC37BB4DF}
  [127] = {link=FB88829F-F043-4942-9C93-D2BA50858194}
public dio _dOutUser[96]
  [32] = {link=FastIO\fOut0}
  [33] = {link=FastIO\fOut1}
public dio dInAckAlarmCmd = {link=DB25555B-9639-404C-BF41-A1E4182E7853}
public dio dInEndCmd = {link=0D6C59A5-572E-4845-9D24-D0618D782DD4}
public dio dInGohomeCmd = {link=A68ADCD7-077C-45ED-AE36-CA1771248567}
public dio dInHoldCmd = {link=F299EF97-EDDD-4BB8-AA07-719E60051D06}
public dio dInPowerOffCmd = {link=1B720B0E-A94A-4B35-8241-512C8CFE7420}
public dio dInPowerOnCmd = {link=1A1317E2-9651-45BA-ACEA-D1820BFA9703}
public dio dInReadJob
public dio dInResetCmd = {link=801699AD-0D4E-40AF-A7AF-E7C40311637E}
public dio dInResetIOCmd = {link=6F68113A-0DD2-4F74-B0DE-02F63C641B3D}
public dio dInStartCmd = {link=842E3CE8-5982-430F-AA8E-B2F701DC178B}
public dio dInStopCmd = {link=CC171C2B-47CE-4C45-9659-7FCDC013CE94}
public dio dInVirtual[128]
  [0] = {link=VirtualIOBoards\VirtualBoard0\%I0}
  [1] = {link=VirtualIOBoards\VirtualBoard0\%I1}
  [2] = {link=VirtualIOBoards\VirtualBoard0\%I2}
  [3] = {link=VirtualIOBoards\VirtualBoard0\%I3}
  [4] = {link=VirtualIOBoards\VirtualBoard0\%I4}
  [5] = {link=VirtualIOBoards\VirtualBoard0\%I5}
  [6] = {link=VirtualIOBoards\VirtualBoard0\%I6}
  [7] = {link=VirtualIOBoards\VirtualBoard0\%I7}
  [8] = {link=VirtualIOBoards\VirtualBoard0\%I8}
  [9] = {link=VirtualIOBoards\VirtualBoard0\%I9}
  [10] = {link=VirtualIOBoards\VirtualBoard0\%I10}
  [11] = {link=VirtualIOBoards\VirtualBoard0\%I11}
  [12] = {link=VirtualIOBoards\VirtualBoard0\%I12}
  [13] = {link=VirtualIOBoards\VirtualBoard0\%I13}
  [14] = {link=VirtualIOBoards\VirtualBoard0\%I14}
  [15] = {link=VirtualIOBoards\VirtualBoard0\%I15}
  [16] = {link=VirtualIOBoards\VirtualBoard0\%I16}
  [17] = {link=VirtualIOBoards\VirtualBoard0\%I17}
  [18] = {link=VirtualIOBoards\VirtualBoard0\%I18}
  [19] = {link=VirtualIOBoards\VirtualBoard0\%I19}
  [20] = {link=VirtualIOBoards\VirtualBoard0\%I20}
  [21] = {link=VirtualIOBoards\VirtualBoard0\%I21}
  [22] = {link=VirtualIOBoards\VirtualBoard0\%I22}
  [23] = {link=VirtualIOBoards\VirtualBoard0\%I23}
  [24] = {link=VirtualIOBoards\VirtualBoard0\%I24}
  [25] = {link=VirtualIOBoards\VirtualBoard0\%I25}
  [26] = {link=VirtualIOBoards\VirtualBoard0\%I26}
  [27] = {link=VirtualIOBoards\VirtualBoard0\%I27}
  [28] = {link=VirtualIOBoards\VirtualBoard0\%I28}
  [29] = {link=VirtualIOBoards\VirtualBoard0\%I29}
  [30] = {link=VirtualIOBoards\VirtualBoard0\%I30}
  [31] = {link=VirtualIOBoards\VirtualBoard0\%I31}
  [32] = {link=VirtualIOBoards\VirtualBoard0\%I32}
  [33] = {link=VirtualIOBoards\VirtualBoard0\%I33}
  [34] = {link=VirtualIOBoards\VirtualBoard0\%I34}
  [35] = {link=VirtualIOBoards\VirtualBoard0\%I35}
  [36] = {link=VirtualIOBoards\VirtualBoard0\%I36}
  [37] = {link=VirtualIOBoards\VirtualBoard0\%I37}
  [38] = {link=VirtualIOBoards\VirtualBoard0\%I38}
  [39] = {link=VirtualIOBoards\VirtualBoard0\%I39}
  [40] = {link=VirtualIOBoards\VirtualBoard0\%I40}
  [41] = {link=VirtualIOBoards\VirtualBoard0\%I41}
  [42] = {link=VirtualIOBoards\VirtualBoard0\%I42}
  [43] = {link=VirtualIOBoards\VirtualBoard0\%I43}
  [44] = {link=VirtualIOBoards\VirtualBoard0\%I44}
  [45] = {link=VirtualIOBoards\VirtualBoard0\%I45}
  [46] = {link=VirtualIOBoards\VirtualBoard0\%I46}
  [47] = {link=VirtualIOBoards\VirtualBoard0\%I47}
  [48] = {link=VirtualIOBoards\VirtualBoard0\%I48}
  [49] = {link=VirtualIOBoards\VirtualBoard0\%I49}
  [50] = {link=VirtualIOBoards\VirtualBoard0\%I50}
  [51] = {link=VirtualIOBoards\VirtualBoard0\%I51}
  [52] = {link=VirtualIOBoards\VirtualBoard0\%I52}
  [53] = {link=VirtualIOBoards\VirtualBoard0\%I53}
  [54] = {link=VirtualIOBoards\VirtualBoard0\%I54}
  [55] = {link=VirtualIOBoards\VirtualBoard0\%I55}
  [56] = {link=VirtualIOBoards\VirtualBoard0\%I56}
  [57] = {link=VirtualIOBoards\VirtualBoard0\%I57}
  [58] = {link=VirtualIOBoards\VirtualBoard0\%I58}
  [59] = {link=VirtualIOBoards\VirtualBoard0\%I59}
  [60] = {link=VirtualIOBoards\VirtualBoard0\%I60}
  [61] = {link=VirtualIOBoards\VirtualBoard0\%I61}
  [62] = {link=VirtualIOBoards\VirtualBoard0\%I62}
  [63] = {link=VirtualIOBoards\VirtualBoard0\%I63}
  [64] = {link=VirtualIOBoards\VirtualBoard0\%I64}
  [65] = {link=VirtualIOBoards\VirtualBoard0\%I65}
  [66] = {link=VirtualIOBoards\VirtualBoard0\%I66}
  [67] = {link=VirtualIOBoards\VirtualBoard0\%I67}
  [68] = {link=VirtualIOBoards\VirtualBoard0\%I68}
  [69] = {link=VirtualIOBoards\VirtualBoard0\%I69}
  [70] = {link=VirtualIOBoards\VirtualBoard0\%I70}
  [71] = {link=VirtualIOBoards\VirtualBoard0\%I71}
  [72] = {link=VirtualIOBoards\VirtualBoard0\%I72}
  [73] = {link=VirtualIOBoards\VirtualBoard0\%I73}
  [74] = {link=VirtualIOBoards\VirtualBoard0\%I74}
  [75] = {link=VirtualIOBoards\VirtualBoard0\%I75}
  [76] = {link=VirtualIOBoards\VirtualBoard0\%I76}
  [77] = {link=VirtualIOBoards\VirtualBoard0\%I77}
  [78] = {link=VirtualIOBoards\VirtualBoard0\%I78}
  [79] = {link=VirtualIOBoards\VirtualBoard0\%I79}
  [80] = {link=VirtualIOBoards\VirtualBoard0\%I80}
  [81] = {link=VirtualIOBoards\VirtualBoard0\%I81}
  [82] = {link=VirtualIOBoards\VirtualBoard0\%I82}
  [83] = {link=VirtualIOBoards\VirtualBoard0\%I83}
  [84] = {link=VirtualIOBoards\VirtualBoard0\%I84}
  [85] = {link=VirtualIOBoards\VirtualBoard0\%I85}
  [86] = {link=VirtualIOBoards\VirtualBoard0\%I86}
  [87] = {link=VirtualIOBoards\VirtualBoard0\%I87}
  [88] = {link=VirtualIOBoards\VirtualBoard0\%I88}
  [89] = {link=VirtualIOBoards\VirtualBoard0\%I89}
  [90] = {link=VirtualIOBoards\VirtualBoard0\%I90}
  [91] = {link=VirtualIOBoards\VirtualBoard0\%I91}
  [92] = {link=VirtualIOBoards\VirtualBoard0\%I92}
  [93] = {link=VirtualIOBoards\VirtualBoard0\%I93}
  [94] = {link=VirtualIOBoards\VirtualBoard0\%I94}
  [95] = {link=VirtualIOBoards\VirtualBoard0\%I95}
  [96] = {link=VirtualIOBoards\VirtualBoard0\%I96}
  [97] = {link=VirtualIOBoards\VirtualBoard0\%I97}
  [98] = {link=VirtualIOBoards\VirtualBoard0\%I98}
  [99] = {link=VirtualIOBoards\VirtualBoard0\%I99}
  [100] = {link=VirtualIOBoards\VirtualBoard0\%I100}
  [101] = {link=VirtualIOBoards\VirtualBoard0\%I101}
  [102] = {link=VirtualIOBoards\VirtualBoard0\%I102}
  [103] = {link=VirtualIOBoards\VirtualBoard0\%I103}
  [104] = {link=VirtualIOBoards\VirtualBoard0\%I104}
  [105] = {link=VirtualIOBoards\VirtualBoard0\%I105}
  [106] = {link=VirtualIOBoards\VirtualBoard0\%I106}
  [107] = {link=VirtualIOBoards\VirtualBoard0\%I107}
  [108] = {link=VirtualIOBoards\VirtualBoard0\%I108}
  [109] = {link=VirtualIOBoards\VirtualBoard0\%I109}
  [110] = {link=VirtualIOBoards\VirtualBoard0\%I110}
  [111] = {link=VirtualIOBoards\VirtualBoard0\%I111}
  [112] = {link=VirtualIOBoards\VirtualBoard0\%I112}
  [113] = {link=VirtualIOBoards\VirtualBoard0\%I113}
  [114] = {link=VirtualIOBoards\VirtualBoard0\%I114}
  [115] = {link=VirtualIOBoards\VirtualBoard0\%I115}
  [116] = {link=VirtualIOBoards\VirtualBoard0\%I116}
  [117] = {link=VirtualIOBoards\VirtualBoard0\%I117}
  [118] = {link=VirtualIOBoards\VirtualBoard0\%I118}
  [119] = {link=VirtualIOBoards\VirtualBoard0\%I119}
  [120] = {link=VirtualIOBoards\VirtualBoard0\%I120}
  [121] = {link=VirtualIOBoards\VirtualBoard0\%I121}
  [122] = {link=VirtualIOBoards\VirtualBoard0\%I122}
  [123] = {link=VirtualIOBoards\VirtualBoard0\%I123}
  [124] = {link=VirtualIOBoards\VirtualBoard0\%I124}
  [125] = {link=VirtualIOBoards\VirtualBoard0\%I125}
  [126] = {link=VirtualIOBoards\VirtualBoard0\%I126}
  [127] = {link=VirtualIOBoards\VirtualBoard0\%I127}
public dio dInput[128]
  [0] = {link=801699AD-0D4E-40AF-A7AF-E7C40311637E}
  [1] = {link=842E3CE8-5982-430F-AA8E-B2F701DC178B}
  [2] = {link=F299EF97-EDDD-4BB8-AA07-719E60051D06}
  [3] = {link=0D6C59A5-572E-4845-9D24-D0618D782DD4}
  [4] = {link=CC171C2B-47CE-4C45-9659-7FCDC013CE94}
  [5] = {link=1A1317E2-9651-45BA-ACEA-D1820BFA9703}
  [6] = {link=1B720B0E-A94A-4B35-8241-512C8CFE7420}
  [7] = {link=6F68113A-0DD2-4F74-B0DE-02F63C641B3D}
  [8] = {link=DB25555B-9639-404C-BF41-A1E4182E7853}
  [9] = {link=A68ADCD7-077C-45ED-AE36-CA1771248567}
  [10] = {link=3971923C-046E-4FB8-8CDF-8298982DD00B}
  [11] = {link=C253DB67-AB15-493D-BA5F-F7404DA89E40}
  [12] = {link=5F58F424-9E7E-46E6-B5AD-37E850D30CCF}
  [13] = {link=0B266260-B4AD-4902-9CA8-DAC05E19210B}
  [14] = {link=20B44CE4-2E83-403B-A39C-4F8E5CA01265}
  [15] = {link=CD23C02B-CC02-4E28-82D0-6EB1534712A8}
  [16] = {link=550C0093-735F-4929-AB88-92E210EEA585}
  [17] = {link=58675BC9-A902-44A6-9D1E-CDCDD371E5BF}
  [18] = {link=C6C06F3F-E54C-4EE8-B5A1-0B392CB95D19}
  [19] = {link=E7996F97-FFB6-4A1D-8389-FC391F807530}
  [20] = {link=545E5659-957E-409A-983D-845A312BF10F}
  [21] = {link=896C2D61-98DD-43B3-A9FF-B63B82E13F66}
  [22] = {link=CB058ED0-A460-493F-ACD8-83515F19CB22}
  [23] = {link=8EC8BEC8-3882-4E09-82EB-ED6F4043F345}
  [24] = {link=6614FE1F-5D84-418F-8C43-3AD6E08D9885}
  [25] = {link=A0D729AE-192B-4443-98B3-A6978F97C45B}
  [26] = {link=8274EAD0-4711-40CE-9532-B3E4F6D5E848}
  [27] = {link=A4D7A453-0050-4322-BCBB-255C4251B0BA}
  [28] = {link=0CFB91EB-8B07-41BC-89A1-F8BBECCF0624}
  [29] = {link=4F7299CD-79A3-4FE2-8435-19083E83C2B9}
  [30] = {link=E49B7D09-65F8-4955-B810-3C508C434830}
  [31] = {link=2BAB1321-D2BB-48C2-8DEA-1230FF1A9D85}
  [32] = {link=C00D5C02-BF78-4EF5-B868-C5B31E42BE7F}
  [33] = {link=96859C69-E3EF-4F26-913D-E25096C13C5F}
  [34] = {link=7920EEE9-3DBF-43F3-9541-7FBE207ECE53}
  [35] = {link=1DB9160A-F63F-4C13-93B5-492FEDD177E2}
  [36] = {link=1FC4D9B1-EE44-4A9B-A22D-5889BB08EE1E}
  [37] = {link=BF970AFE-565C-4857-97A6-5A54DDAE79B6}
  [38] = {link=F909C748-B7A8-4470-A6FD-BA1A46FE4E68}
  [39] = {link=8517CD21-2BAD-4F53-9136-89235F4060C6}
  [40] = {link=6DDBB7AB-AC7B-4F3D-A091-1238925E0448}
  [41] = {link=C3CF7374-59EF-4029-99B4-FC98E25808BB}
  [42] = {link=90C02E77-8235-444D-99EB-D816EF90AFE5}
  [43] = {link=E44556E2-741A-40A0-89B2-8E32677B3EB1}
  [44] = {link=D8AFCC23-6F61-4ADD-8DE3-3FE1547AD28D}
  [45] = {link=98BC2888-38BC-4A33-A762-BDEC3E36173F}
  [46] = {link=A24DA26D-2F10-46AE-809B-0B04336865AA}
  [47] = {link=04D21FA2-EBE1-4E66-8338-7CB17174A724}
  [48] = {link=E766472B-9569-4911-A858-6F7708718D01}
  [49] = {link=92C360C1-157E-40E1-9184-03D53ECDF3F7}
  [50] = {link=6E33B145-BAC8-48E7-A184-E5A9D90B515B}
  [51] = {link=D5FDB290-CB76-4852-8AF4-F9B6FA5D3E2D}
  [52] = {link=547C3630-B2EA-42F8-AB37-EEB4C81AA149}
  [53] = {link=A60C469C-4F75-4C30-9347-66365041DE79}
  [54] = {link=6E14BCEF-8B69-4038-B259-0EF712D2AB66}
  [55] = {link=B19F0E1B-CE25-49C3-9ED7-92404708DBC9}
  [56] = {link=AFC49D6D-7F53-41F5-8159-6058E9291542}
  [57] = {link=BB08126F-937C-4C50-9A1C-252CB13BB25C}
  [58] = {link=15BF4171-EFAA-47B7-BEF9-A698BE11011C}
  [59] = {link=9A261803-1F52-41D2-8355-1C79BF1BB94D}
  [60] = {link=18F63136-91BD-4FEE-8DA3-2AA9D2E8FFA8}
  [61] = {link=55E89D2C-C808-4026-99D2-85E324C475F9}
  [62] = {link=45535323-0512-46DB-8EB0-4BF3F55D73C7}
  [63] = {link=23943399-CEE5-49D9-BFD9-55B5920F548B}
  [64] = {link=364F41EB-6BA1-4700-BD0A-C2236839044E}
  [65] = {link=96EFCAAE-6B9A-4070-B9EC-2035BA94CCB3}
  [66] = {link=FD79DB68-803F-47E7-8305-8CFFFE519C88}
  [67] = {link=82CF98E3-5511-4523-9501-B4BBAD9DC96D}
  [68] = {link=43A446B7-3C25-4DD5-9597-27365DBE2539}
  [69] = {link=01367322-9745-4163-BFB8-DF881D521F4A}
  [70] = {link=1F635259-38C5-4AB2-B093-ADA4F82FD92B}
  [71] = {link=80065B3A-E7EF-4B6D-A30A-AC2F8A1FF9BD}
  [72] = {link=138692BF-FCCE-4B34-B0E8-8C4B22C67F12}
  [73] = {link=2F598E66-6704-43A6-A433-14D902C15D10}
  [74] = {link=3D7C9642-411B-40D3-B3B9-C83D24259AF4}
  [75] = {link=2E14C0AE-1F04-4256-8959-DEAD28BB69AE}
  [76] = {link=D90512A1-D0E1-41B2-8294-59D7C1ADD8E0}
  [77] = {link=F9EFA2A2-C655-4B55-8F3F-AAE77A6FD751}
  [78] = {link=8C43F822-1313-4C63-84D2-76D62B96A58F}
  [79] = {link=0BE51982-5E8E-4776-A637-0836608FA4D4}
  [80] = {link=5CC26A0C-A759-4F9D-9C90-7643106A4280}
  [81] = {link=6B2348DB-D0C3-44B1-96EA-09FBC0D6D1F3}
  [82] = {link=091DC27E-E2EB-463E-8E4B-08B48E663650}
  [83] = {link=EC5520D5-F711-48B3-AE90-97344DDBEE5C}
  [84] = {link=E02811C8-C36E-4E92-B28C-81A727813C5B}
  [85] = {link=39EB69C5-9612-415D-9A77-D013E3B8CFD4}
  [86] = {link=FD4FFC3C-593A-4304-8BB2-18534DB95237}
  [87] = {link=D2ECCFF1-C6D1-48A4-B3A9-F333711A9798}
  [88] = {link=13EA7043-3380-41E5-9177-AAC787C21C39}
  [89] = {link=5475660F-31B7-47C3-808C-FBAB066EFE6D}
  [90] = {link=93D7CC16-1244-4B9F-85C2-564B516A38A6}
  [91] = {link=A2A5B44E-CAC8-47F1-A810-875EED5095FB}
  [92] = {link=2F9951E4-3414-412E-A45B-55B5D632DA1B}
  [93] = {link=916866A1-8E9C-42B7-A695-7CB9D795E148}
  [94] = {link=CA3200CB-BA9D-4435-B593-6CDDBB86F10C}
  [95] = {link=49AC3AF5-F49B-42A1-90B2-5DB7D6C7E051}
  [96] = {link=64E7B72A-8AE1-43E7-9A21-FF4DABD03910}
  [97] = {link=7BA0757A-43B7-4994-86FC-1740DE8C159E}
  [98] = {link=5ACF5B88-9BD6-435A-8F3F-752FE88E7935}
  [99] = {link=70DFB9C6-9CA4-44C9-8464-A31BA0D039F5}
  [100] = {link=55D5D0F9-E23A-40DA-9955-6BCB63B37099}
  [101] = {link=1AB52030-AE2C-417B-9C38-1633EF57A0DB}
  [102] = {link=FFE2E20E-ABB5-4A36-BE3B-E714CB40E85A}
  [103] = {link=83BC89DD-B780-47A7-BBF0-017BDC2BA365}
  [104] = {link=10D6F5C6-79FE-4371-9CC9-A814346F77C1}
  [105] = {link=240957B0-B56A-4DFB-9281-23480961F3F1}
  [106] = {link=92C2EE73-BB65-4A97-8029-77FB60FFC23C}
  [107] = {link=62C2F98E-E7EB-49ED-971A-83A5444F6152}
  [108] = {link=58CC62E1-4595-401C-8E2F-3122D818CC74}
  [109] = {link=6D2EBC96-6FF5-40C1-83D6-CC8DD3D9FC3A}
  [110] = {link=AEC5DD07-0ABE-4FC2-A89A-ED52FEBBCAD7}
  [111] = {link=D289FF49-1CD8-4174-B7A5-8E375EB48B35}
  [112] = {link=4D3459D2-B2AE-4602-8654-6AD44AA154CE}
  [113] = {link=BE4318FA-0CA3-4B50-ACFD-D0BD90E002BB}
  [114] = {link=03734564-3942-45B2-807F-C861E4A00B4D}
  [115] = {link=18C4B14F-9C0F-4159-B56F-314AFF4BFABC}
  [116] = {link=A703F976-FEB8-4965-8F5A-CAD8585E54F7}
  [117] = {link=F3814F6C-1F81-45E4-8DE4-AB9F0C1AC9C1}
  [118] = {link=CD215C83-5C8C-4339-BF6C-DDE6EDBF5021}
  [119] = {link=295A35FF-B8CC-4A25-BC99-5CC4EFE79E3D}
  [120] = {link=7D822E1A-7C34-46E1-A06C-E10F3FD6B4DE}
  [121] = {link=4A23737B-5C9C-4372-A68A-8F60451AD439}
  [122] = {link=B2909A16-C926-42A5-8387-168FB9DA6D2A}
  [123] = {link=36FA5061-3D34-4793-BCBA-E09767B9821D}
  [124] = {link=0AE8B5A8-7356-480B-AAA1-20AFD496F398}
  [125] = {link=DB043A0E-80EF-4F10-9CBC-7A049A7AEFDE}
  [126] = {link=951CF18F-CA29-47EF-A085-39A8D6CD28C1}
  [127] = {link=6FC2F7D5-08CF-47CC-86FA-1AC31B966FFD}
public dio dOGohomeing = {link=75D4F3C1-C356-4EDA-B423-02C90835EA7D}
public dio dOMcpEstop = {link=C4522756-21A9-4D8A-B398-209F6EFB0977}
public dio dORbAlarm = {link=07A4EEA8-4CAE-47C3-9487-42EFEC0C0C8E}
public dio dORbAtHome = {link=3F319035-E82A-4D07-9742-3AFC501B53DF}
public dio dORbAutoMode = {link=16CB4CF9-3A13-4F09-B6E9-D967DFB15E25}
public dio dORbEnable = {link=698A0489-9B90-43A7-B0CD-777095A36007}
public dio dORbEstop = {link=VirtualIOBoards\VirtualBoard0\%Q13}
public dio dORbHeartbeat = {link=2087A18A-21B3-4E9A-90F0-0A72D013BBC2}
public dio dORbHeld = {link=79705501-C546-4790-A460-3F340ADFDE5C}
public dio dORbManualMode = {link=734EBAF3-2CA8-4D3F-A8BB-E168C1322725}
public dio dORbMoving = {link=93BF17B5-5C7E-43C6-9C42-3B6025772815}
public dio dORbPowerOn = {link=1CC4B59E-3D71-495F-A34B-473B0A37D044}
public dio dORbReady = {link=364EC08F-C077-495B-A954-158507D3C26C}
public dio dORbRunning = {link=289A5E8D-11F3-4BEB-8FA4-200735E3A2B7}
public dio dORbStopped = {link=813E3F4B-A1DE-4C5D-8EAB-0242B6D8A546}
public dio dORbTaskRunOk = {link=63159677-63A9-4936-A8C6-E65B2885D59F}
public dio dOutVirtual[128]
  [0] = {link=VirtualIOBoards\VirtualBoard0\%Q0}
  [1] = {link=VirtualIOBoards\VirtualBoard0\%Q1}
  [2] = {link=VirtualIOBoards\VirtualBoard0\%Q2}
  [3] = {link=VirtualIOBoards\VirtualBoard0\%Q3}
  [4] = {link=VirtualIOBoards\VirtualBoard0\%Q4}
  [5] = {link=VirtualIOBoards\VirtualBoard0\%Q5}
  [6] = {link=VirtualIOBoards\VirtualBoard0\%Q6}
  [7] = {link=VirtualIOBoards\VirtualBoard0\%Q7}
  [8] = {link=VirtualIOBoards\VirtualBoard0\%Q8}
  [9] = {link=VirtualIOBoards\VirtualBoard0\%Q9}
  [10] = {link=VirtualIOBoards\VirtualBoard0\%Q10}
  [11] = {link=VirtualIOBoards\VirtualBoard0\%Q11}
  [12] = {link=VirtualIOBoards\VirtualBoard0\%Q12}
  [13] = {link=VirtualIOBoards\VirtualBoard0\%Q13}
  [14] = {link=VirtualIOBoards\VirtualBoard0\%Q14}
  [15] = {link=VirtualIOBoards\VirtualBoard0\%Q15}
  [16] = {link=VirtualIOBoards\VirtualBoard0\%Q16}
  [17] = {link=VirtualIOBoards\VirtualBoard0\%Q17}
  [18] = {link=VirtualIOBoards\VirtualBoard0\%Q18}
  [19] = {link=VirtualIOBoards\VirtualBoard0\%Q19}
  [20] = {link=VirtualIOBoards\VirtualBoard0\%Q20}
  [21] = {link=VirtualIOBoards\VirtualBoard0\%Q21}
  [22] = {link=VirtualIOBoards\VirtualBoard0\%Q22}
  [23] = {link=VirtualIOBoards\VirtualBoard0\%Q23}
  [24] = {link=VirtualIOBoards\VirtualBoard0\%Q24}
  [25] = {link=VirtualIOBoards\VirtualBoard0\%Q25}
  [26] = {link=VirtualIOBoards\VirtualBoard0\%Q26}
  [27] = {link=VirtualIOBoards\VirtualBoard0\%Q27}
  [28] = {link=VirtualIOBoards\VirtualBoard0\%Q28}
  [29] = {link=VirtualIOBoards\VirtualBoard0\%Q29}
  [30] = {link=VirtualIOBoards\VirtualBoard0\%Q30}
  [31] = {link=VirtualIOBoards\VirtualBoard0\%Q31}
  [32] = {link=VirtualIOBoards\VirtualBoard0\%Q32}
  [33] = {link=VirtualIOBoards\VirtualBoard0\%Q33}
  [34] = {link=VirtualIOBoards\VirtualBoard0\%Q34}
  [35] = {link=VirtualIOBoards\VirtualBoard0\%Q35}
  [36] = {link=VirtualIOBoards\VirtualBoard0\%Q36}
  [37] = {link=VirtualIOBoards\VirtualBoard0\%Q37}
  [38] = {link=VirtualIOBoards\VirtualBoard0\%Q38}
  [39] = {link=VirtualIOBoards\VirtualBoard0\%Q39}
  [40] = {link=VirtualIOBoards\VirtualBoard0\%Q40}
  [41] = {link=VirtualIOBoards\VirtualBoard0\%Q41}
  [42] = {link=VirtualIOBoards\VirtualBoard0\%Q42}
  [43] = {link=VirtualIOBoards\VirtualBoard0\%Q43}
  [44] = {link=VirtualIOBoards\VirtualBoard0\%Q44}
  [45] = {link=VirtualIOBoards\VirtualBoard0\%Q45}
  [46] = {link=VirtualIOBoards\VirtualBoard0\%Q46}
  [47] = {link=VirtualIOBoards\VirtualBoard0\%Q47}
  [48] = {link=VirtualIOBoards\VirtualBoard0\%Q48}
  [49] = {link=VirtualIOBoards\VirtualBoard0\%Q49}
  [50] = {link=VirtualIOBoards\VirtualBoard0\%Q50}
  [51] = {link=VirtualIOBoards\VirtualBoard0\%Q51}
  [52] = {link=VirtualIOBoards\VirtualBoard0\%Q52}
  [53] = {link=VirtualIOBoards\VirtualBoard0\%Q53}
  [54] = {link=VirtualIOBoards\VirtualBoard0\%Q54}
  [55] = {link=VirtualIOBoards\VirtualBoard0\%Q55}
  [56] = {link=VirtualIOBoards\VirtualBoard0\%Q56}
  [57] = {link=VirtualIOBoards\VirtualBoard0\%Q57}
  [58] = {link=VirtualIOBoards\VirtualBoard0\%Q58}
  [59] = {link=VirtualIOBoards\VirtualBoard0\%Q59}
  [60] = {link=VirtualIOBoards\VirtualBoard0\%Q60}
  [61] = {link=VirtualIOBoards\VirtualBoard0\%Q61}
  [62] = {link=VirtualIOBoards\VirtualBoard0\%Q62}
  [63] = {link=VirtualIOBoards\VirtualBoard0\%Q63}
  [64] = {link=VirtualIOBoards\VirtualBoard0\%Q64}
  [65] = {link=VirtualIOBoards\VirtualBoard0\%Q65}
  [66] = {link=VirtualIOBoards\VirtualBoard0\%Q66}
  [67] = {link=VirtualIOBoards\VirtualBoard0\%Q67}
  [68] = {link=VirtualIOBoards\VirtualBoard0\%Q68}
  [69] = {link=VirtualIOBoards\VirtualBoard0\%Q69}
  [70] = {link=VirtualIOBoards\VirtualBoard0\%Q70}
  [71] = {link=VirtualIOBoards\VirtualBoard0\%Q71}
  [72] = {link=VirtualIOBoards\VirtualBoard0\%Q72}
  [73] = {link=VirtualIOBoards\VirtualBoard0\%Q73}
  [74] = {link=VirtualIOBoards\VirtualBoard0\%Q74}
  [75] = {link=VirtualIOBoards\VirtualBoard0\%Q75}
  [76] = {link=VirtualIOBoards\VirtualBoard0\%Q76}
  [77] = {link=VirtualIOBoards\VirtualBoard0\%Q77}
  [78] = {link=VirtualIOBoards\VirtualBoard0\%Q78}
  [79] = {link=VirtualIOBoards\VirtualBoard0\%Q79}
  [80] = {link=VirtualIOBoards\VirtualBoard0\%Q80}
  [81] = {link=VirtualIOBoards\VirtualBoard0\%Q81}
  [82] = {link=VirtualIOBoards\VirtualBoard0\%Q82}
  [83] = {link=VirtualIOBoards\VirtualBoard0\%Q83}
  [84] = {link=VirtualIOBoards\VirtualBoard0\%Q84}
  [85] = {link=VirtualIOBoards\VirtualBoard0\%Q85}
  [86] = {link=VirtualIOBoards\VirtualBoard0\%Q86}
  [87] = {link=VirtualIOBoards\VirtualBoard0\%Q87}
  [88] = {link=VirtualIOBoards\VirtualBoard0\%Q88}
  [89] = {link=VirtualIOBoards\VirtualBoard0\%Q89}
  [90] = {link=VirtualIOBoards\VirtualBoard0\%Q90}
  [91] = {link=VirtualIOBoards\VirtualBoard0\%Q91}
  [92] = {link=VirtualIOBoards\VirtualBoard0\%Q92}
  [93] = {link=VirtualIOBoards\VirtualBoard0\%Q93}
  [94] = {link=VirtualIOBoards\VirtualBoard0\%Q94}
  [95] = {link=VirtualIOBoards\VirtualBoard0\%Q95}
  [96] = {link=VirtualIOBoards\VirtualBoard0\%Q96}
  [97] = {link=VirtualIOBoards\VirtualBoard0\%Q97}
  [98] = {link=VirtualIOBoards\VirtualBoard0\%Q98}
  [99] = {link=VirtualIOBoards\VirtualBoard0\%Q99}
  [100] = {link=VirtualIOBoards\VirtualBoard0\%Q100}
  [101] = {link=VirtualIOBoards\VirtualBoard0\%Q101}
  [102] = {link=VirtualIOBoards\VirtualBoard0\%Q102}
  [103] = {link=VirtualIOBoards\VirtualBoard0\%Q103}
  [104] = {link=VirtualIOBoards\VirtualBoard0\%Q104}
  [105] = {link=VirtualIOBoards\VirtualBoard0\%Q105}
  [106] = {link=VirtualIOBoards\VirtualBoard0\%Q106}
  [107] = {link=VirtualIOBoards\VirtualBoard0\%Q107}
  [108] = {link=VirtualIOBoards\VirtualBoard0\%Q108}
  [109] = {link=VirtualIOBoards\VirtualBoard0\%Q109}
  [110] = {link=VirtualIOBoards\VirtualBoard0\%Q110}
  [111] = {link=VirtualIOBoards\VirtualBoard0\%Q111}
  [112] = {link=VirtualIOBoards\VirtualBoard0\%Q112}
  [113] = {link=VirtualIOBoards\VirtualBoard0\%Q113}
  [114] = {link=VirtualIOBoards\VirtualBoard0\%Q114}
  [115] = {link=VirtualIOBoards\VirtualBoard0\%Q115}
  [116] = {link=VirtualIOBoards\VirtualBoard0\%Q116}
  [117] = {link=VirtualIOBoards\VirtualBoard0\%Q117}
  [118] = {link=VirtualIOBoards\VirtualBoard0\%Q118}
  [119] = {link=VirtualIOBoards\VirtualBoard0\%Q119}
  [120] = {link=VirtualIOBoards\VirtualBoard0\%Q120}
  [121] = {link=VirtualIOBoards\VirtualBoard0\%Q121}
  [122] = {link=VirtualIOBoards\VirtualBoard0\%Q122}
  [123] = {link=VirtualIOBoards\VirtualBoard0\%Q123}
  [124] = {link=VirtualIOBoards\VirtualBoard0\%Q124}
  [125] = {link=VirtualIOBoards\VirtualBoard0\%Q125}
  [126] = {link=VirtualIOBoards\VirtualBoard0\%Q126}
  [127] = {link=VirtualIOBoards\VirtualBoard0\%Q127}
public dio dOutput[128]
  [0] = {link=813E3F4B-A1DE-4C5D-8EAB-0242B6D8A546}
  [1] = {link=364EC08F-C077-495B-A954-158507D3C26C}
  [2] = {link=289A5E8D-11F3-4BEB-8FA4-200735E3A2B7}
  [3] = {link=79705501-C546-4790-A460-3F340ADFDE5C}
  [4] = {link=75D4F3C1-C356-4EDA-B423-02C90835EA7D}
  [5] = {link=3F319035-E82A-4D07-9742-3AFC501B53DF}
  [6] = {link=1CC4B59E-3D71-495F-A34B-473B0A37D044}
  [7] = {link=2087A18A-21B3-4E9A-90F0-0A72D013BBC2}
  [8] = {link=93BF17B5-5C7E-43C6-9C42-3B6025772815}
  [9] = {link=16CB4CF9-3A13-4F09-B6E9-D967DFB15E25}
  [10] = {link=734EBAF3-2CA8-4D3F-A8BB-E168C1322725}
  [11] = {link=07A4EEA8-4CAE-47C3-9487-42EFEC0C0C8E}
  [12] = {link=63159677-63A9-4936-A8C6-E65B2885D59F}
  [13] = {link=698A0489-9B90-43A7-B0CD-777095A36007}
  [14] = {link=C4522756-21A9-4D8A-B398-209F6EFB0977}
  [15] = {link=E3974102-9CCD-497B-BD29-7D9DDF1F0662}
  [16] = {link=D7E9BDA6-AD73-4469-BD4D-C9D8F1711105}
  [17] = {link=C0E9CDD3-3C86-4E8A-BB76-29DD4E724269}
  [18] = {link=19A15CFF-CD59-4687-8101-878C6D297AD0}
  [19] = {link=F886CB4C-7C2D-4AEE-8DA8-19CCB8826A1C}
  [20] = {link=44B2E852-2BDD-46AD-B032-142EDC75806B}
  [21] = {link=E6202C42-8108-4A9C-988A-BA326395584A}
  [22] = {link=4A293BE2-BE94-462E-ACFA-7E01BA496DDB}
  [23] = {link=C4CC4269-4D2F-4B53-89D1-5B6F0F9E20C5}
  [24] = {link=976E4904-0F44-43DA-867D-0C06FC7F067A}
  [25] = {link=26F2F168-65FE-450B-BE6F-27BCBE8A7C37}
  [26] = {link=58979B7C-3302-40C0-9293-D8BDE318359F}
  [27] = {link=32E62FFE-3CE0-449B-8ADB-B460A9E5DE54}
  [28] = {link=1778E8D0-D57F-4F6E-A6A4-A7E0DC8A5FDF}
  [29] = {link=BB6EEE31-C681-41BA-8160-A41199CEAD02}
  [30] = {link=58577585-C0FF-479D-B4D2-FF8F04E87201}
  [31] = {link=E4789C35-874D-4E09-8AF9-741C03AAD9B4}
  [32] = {link=AB4C11BC-0698-4F05-9F77-33C54B19FD7D}
  [33] = {link=A971CAAA-D369-4C08-BB4B-F444CDC4D2F0}
  [34] = {link=EE574E0A-35B5-4DE1-8C9E-C0DF9CDCDFE6}
  [35] = {link=7532402E-1B90-4BA9-83CA-579B1F726874}
  [36] = {link=6F6C7C8F-8851-47C2-9B8E-D33C24B9D39F}
  [37] = {link=4A5CAAE4-C9CD-4421-94AD-56079246CA39}
  [38] = {link=EB7E2C34-F887-4C3F-97E0-01834D630C5E}
  [39] = {link=BDBB409A-6EC7-4423-9FF9-A638D02BF80E}
  [40] = {link=E136414E-B9B9-4DA1-8541-C1A78F1E80BF}
  [41] = {link=8E4798E6-5BA8-40FC-8B4C-D83695D2AB51}
  [42] = {link=28472F68-DF34-4C50-9023-A219CE2C4B1B}
  [43] = {link=1DB5BD39-DE07-40ED-B700-8C7874B04DB0}
  [44] = {link=88484DFD-5685-4FE3-BD11-1467A80C9B34}
  [45] = {link=2F5F1623-83AA-4A31-A803-F6FA4D4BE14A}
  [46] = {link=519B5132-0D61-4FA5-ABD4-96724AED25E8}
  [47] = {link=661BE778-7099-413C-A47D-EC9A4ECEF23E}
  [48] = {link=53B2124C-FE98-440B-9A3D-84530B55B740}
  [49] = {link=229E980F-A7B4-4859-9EE1-BA541F4B5A16}
  [50] = {link=1FA4F26D-23CC-42E9-A819-02B2DD7006DA}
  [51] = {link=2AEDD394-CA8D-4F24-A299-43D2A058ACD5}
  [52] = {link=C28EB1DF-BACA-4254-A598-B532E330438E}
  [53] = {link=E7F3183B-4DF3-459A-ADF7-79D82988755C}
  [54] = {link=2614E536-799A-40AF-9560-80A760021F62}
  [55] = {link=757B7056-4991-459D-8227-2BCDF4BE047B}
  [56] = {link=8C99F1DA-9DA9-4BDF-B60F-FD54ABC54EFA}
  [57] = {link=5AA809C1-68E1-4A24-9F04-C8074121C64A}
  [58] = {link=4A164529-4FC6-4374-9AB6-7CFCFB13974B}
  [59] = {link=70724C45-B1FB-42FE-A3A2-C0AB8AA81684}
  [60] = {link=9EE71F53-97CD-4882-A49E-A6F1E8BC9441}
  [61] = {link=81277848-FDAC-47B2-B4F0-EFE16B2F5C1C}
  [62] = {link=E56352E6-5F75-449C-AD2C-249D38B077FB}
  [63] = {link=5728C013-0742-4355-8E61-1A03F1F076E6}
  [64] = {link=04B33B81-599B-4BDE-99DF-EEC79DF42297}
  [65] = {link=D5C4F9D4-602E-45CC-A360-A9C8DFC51706}
  [66] = {link=0F23F4DE-A6DC-48A8-BD13-38096E17E4BC}
  [67] = {link=725D593E-3E8C-49B9-A0C8-EC5E7EDBEF47}
  [68] = {link=D80F8BA0-A9D7-467A-84F3-2EF911086F28}
  [69] = {link=290333BB-E8D8-473B-B7DA-1770BF97A3BA}
  [70] = {link=3451ABCB-1CE5-49F5-8053-7E43529834C5}
  [71] = {link=1C486D5A-1AEA-494E-AC84-6CEA9FC0F052}
  [72] = {link=0B5202A6-62EE-4D6C-8E76-4A396B266DA1}
  [73] = {link=07376469-6AEC-4E90-A30D-02A336A51CCF}
  [74] = {link=9C60D734-A29B-44DA-837E-97A014720D64}
  [75] = {link=F6F5CEBA-7A13-4322-B86E-E02B17A52B8C}
  [76] = {link=034F848A-A2B4-4107-BA29-37F2DF0B4836}
  [77] = {link=2D3AB11E-A0E7-43D6-A64B-B19DE4EDCA54}
  [78] = {link=6B87E34F-9D7F-4178-ADAD-CF451768FAD1}
  [79] = {link=0BECC0A6-11C6-443C-B8B7-B823C5449F03}
  [80] = {link=0FAFA963-6C61-46BA-8B8E-FD5D821CED0B}
  [81] = {link=E858B3E5-8FFB-4B3B-9E73-58A45F891801}
  [82] = {link=52490A38-A31A-4D56-AA93-4E3292557F7F}
  [83] = {link=07DE5AAD-9C80-4970-8E40-B99AD098B2C3}
  [84] = {link=E76E3858-8352-4107-BC87-39491D8B651A}
  [85] = {link=2B09FA37-BF2E-4ED9-B53F-09BB42630F57}
  [86] = {link=C0D4BCE7-AA67-4991-AD3B-5583CCFF9A80}
  [87] = {link=BBA329F0-9B99-401C-B2C0-5AA54B82A434}
  [88] = {link=1FF771B4-EE27-450D-A9DB-7E394712BF39}
  [89] = {link=19978664-DA67-4FAE-9478-F6C2FD7BC1A1}
  [90] = {link=B280086E-4E78-4C33-A16A-5103EDFD12BA}
  [91] = {link=66D76411-AF4D-465C-BF45-D26D600CE49D}
  [92] = {link=CF5BF486-B482-4F9A-936E-D7550E22D48F}
  [93] = {link=47EF2689-3337-4012-BAD2-52612379B15C}
  [94] = {link=9BC9630D-0782-4292-B056-6CBDA421EF62}
  [95] = {link=CAFB5CCA-B450-480D-9CAD-A29B903F45A9}
  [96] = {link=DCBA4C7F-A728-4F25-89A5-B6259619A80B}
  [97] = {link=6753AC4A-51FA-413E-B4B2-137174F0D507}
  [98] = {link=81370562-9275-47C1-93C0-CB31297CDD20}
  [99] = {link=E6DCC6F0-C964-47CD-B4D7-1BD8BFDA33AE}
  [100] = {link=18C334B4-AE06-448E-96BF-3CD280A2541B}
  [101] = {link=15B48D0D-C668-47AF-A704-10BA0ED6FFE7}
  [102] = {link=DA2930BB-B07C-4C38-ADBB-0FDC55ECF2BB}
  [103] = {link=8DDD8F2E-B5A8-4F54-BD1B-48D04A96C878}
  [104] = {link=72245E17-FF99-4704-8474-EDB79B027BF9}
  [105] = {link=BCF85E34-592F-4BA5-AE76-F1E8F2FD96C1}
  [106] = {link=9ED9CFBB-1644-41A9-955E-D6E7EB6EF2F1}
  [107] = {link=5A6FDD52-29C6-40B7-B97D-88DE84ED4E53}
  [108] = {link=8E4836F5-8A3D-4937-90E9-0F98CBF16A27}
  [109] = {link=4305B788-10E3-4C38-9835-3E94A9820D41}
  [110] = {link=152B6212-6AC5-4D19-A5F9-C32452DCD0BD}
  [111] = {link=60BD22D0-03A0-4632-85E7-7AB9A7B5E9EE}
  [112] = {link=617AC81D-63D2-418A-A221-1A45E82E8F33}
  [113] = {link=DA60158B-5C4B-4C1D-9AEB-3A4C25735862}
  [114] = {link=7E45E59A-6E5F-4DD8-8E87-A62787B5121D}
  [115] = {link=302676B4-AFEF-4A5D-9D0F-7D7EEE15BD09}
  [116] = {link=94FD2E61-B0C4-426E-8CB5-3D13DE4E72D1}
  [117] = {link=5441B2EB-7737-420D-A838-CB6BC6A9AA98}
  [118] = {link=D70A9639-74F8-485B-B1AE-A12B6619BE09}
  [119] = {link=3C4D5DF3-3DD0-4928-9BAC-FF9DB40E9304}
  [120] = {link=389B2383-01D9-4D6D-8093-13CF39736E4D}
  [121] = {link=9C61CF1A-5A0B-480F-A9AF-E365017F4409}
  [122] = {link=D6F4FFC6-5A52-44AE-AAFC-981F5DBD7076}
  [123] = {link=3768B870-3C40-471D-B639-CE39EBCB3865}
  [124] = {link=FCBA4290-2AF9-4EDB-AAB3-C3D5B2BC56ED}
  [125] = {link=FEB8E5C1-4C55-454A-AACA-1D927BE28924}
  [126] = {link=C97B50B1-B825-4E71-A20E-3BFEC37BB4DF}
  [127] = {link=FB88829F-F043-4942-9C93-D2BA50858194}
public dio dRSI9{}
  [RbStop] = {link=Rsi9IO\IusoA1}
  [enabling] = {link=Rsi9IO\Ienabling1}
  [mcpEstop] = {link=Rsi9IO\ImcpEstop1}
public dio dVirtualIO[96]
public dioItem dInItem[128]
  [0]
    dio dDio = {link=801699AD-0D4E-40AF-A7AF-E7C40311637E}
    string sComment = "电机上电"
  [1]
    dio dDio = {link=842E3CE8-5982-430F-AA8E-B2F701DC178B}
    string sComment = "主程序运行"
  [2]
    dio dDio = {link=F299EF97-EDDD-4BB8-AA07-719E60051D06}
    string sComment = "复位报警"
  [3]
    dio dDio = {link=0D6C59A5-572E-4845-9D24-D0618D782DD4}
    string sComment = "PLC系统故障"
  [4]
    dio dDio = {link=CC171C2B-47CE-4C45-9659-7FCDC013CE94}
    string sComment = "备用"
  [5]
    dio dDio = {link=1A1317E2-9651-45BA-ACEA-D1820BFA9703}
    string sComment = "备用"
  [6]
    dio dDio = {link=1B720B0E-A94A-4B35-8241-512C8CFE7420}
    string sComment = "备用"
  [7]
    dio dDio = {link=6F68113A-0DD2-4F74-B0DE-02F63C641B3D}
    string sComment = "备用"
  [8]
    dio dDio = {link=DB25555B-9639-404C-BF41-A1E4182E7853}
    string sComment = "开枪完成"
  [9]
    dio dDio = {link=A68ADCD7-077C-45ED-AE36-CA1771248567}
    string sComment = "关枪完成"
  [10]
    dio dDio = {link=3971923C-046E-4FB8-8CDF-8298982DD00B}
    string sComment = "开始喷涂"
  [11]
    dio dDio = {link=C253DB67-AB15-493D-BA5F-F7404DA89E40}
    string sComment = "备用"
  [12]
    dio dDio = {link=5F58F424-9E7E-46E6-B5AD-37E850D30CCF}
    string sComment = "备用"
  [13]
    dio dDio = {link=0B266260-B4AD-4902-9CA8-DAC05E19210B}
    string sComment = "备用"
  [14]
    dio dDio = {link=20B44CE4-2E83-403B-A39C-4F8E5CA01265}
    string sComment = "备用"
  [15]
    dio dDio = {link=CD23C02B-CC02-4E28-82D0-6EB1534712A8}
    string sComment = "备用"
  [16]
    dio dDio = {link=550C0093-735F-4929-AB88-92E210EEA585}
    string sComment = "备用"
  [17]
    dio dDio = {link=58675BC9-A902-44A6-9D1E-CDCDD371E5BF}
    string sComment = "备用"
  [18]
    dio dDio = {link=C6C06F3F-E54C-4EE8-B5A1-0B392CB95D19}
    string sComment = "备用"
  [19]
    dio dDio = {link=E7996F97-FFB6-4A1D-8389-FC391F807530}
    string sComment = "备用"
  [20]
    dio dDio = {link=545E5659-957E-409A-983D-845A312BF10F}
    string sComment = "备用"
  [21]
    dio dDio = {link=896C2D61-98DD-43B3-A9FF-B63B82E13F66}
    string sComment = "备用"
  [22]
    dio dDio = {link=CB058ED0-A460-493F-ACD8-83515F19CB22}
    string sComment = "备用"
  [23]
    dio dDio = {link=8EC8BEC8-3882-4E09-82EB-ED6F4043F345}
    string sComment = "备用"
  [24]
    dio dDio = {link=6614FE1F-5D84-418F-8C43-3AD6E08D9885}
    string sComment = "备用"
  [25]
    dio dDio = {link=A0D729AE-192B-4443-98B3-A6978F97C45B}
    string sComment = "备用"
  [26]
    dio dDio = {link=8274EAD0-4711-40CE-9532-B3E4F6D5E848}
    string sComment = "备用"
  [27]
    dio dDio = {link=A4D7A453-0050-4322-BCBB-255C4251B0BA}
    string sComment = "备用"
  [28]
    dio dDio = {link=0CFB91EB-8B07-41BC-89A1-F8BBECCF0624}
    string sComment = "备用"
  [29]
    dio dDio = {link=4F7299CD-79A3-4FE2-8435-19083E83C2B9}
    string sComment = "备用"
  [30]
    dio dDio = {link=E49B7D09-65F8-4955-B810-3C508C434830}
    string sComment = "备用"
  [31]
    dio dDio = {link=2BAB1321-D2BB-48C2-8DEA-1230FF1A9D85}
    string sComment = "备用"
  [32]
    dio dDio = {link=C00D5C02-BF78-4EF5-B868-C5B31E42BE7F}
    string sComment = "备用"
  [33]
    dio dDio = {link=96859C69-E3EF-4F26-913D-E25096C13C5F}
    string sComment = "备用"
  [34]
    dio dDio = {link=7920EEE9-3DBF-43F3-9541-7FBE207ECE53}
    string sComment = "备用"
  [35]
    dio dDio = {link=1DB9160A-F63F-4C13-93B5-492FEDD177E2}
    string sComment = "备用"
  [36]
    dio dDio = {link=1FC4D9B1-EE44-4A9B-A22D-5889BB08EE1E}
    string sComment = "备用"
  [37]
    dio dDio = {link=BF970AFE-565C-4857-97A6-5A54DDAE79B6}
    string sComment = "备用"
  [38]
    dio dDio = {link=F909C748-B7A8-4470-A6FD-BA1A46FE4E68}
    string sComment = "备用"
  [39]
    dio dDio = {link=8517CD21-2BAD-4F53-9136-89235F4060C6}
    string sComment = "备用"
  [40]
    dio dDio = {link=6DDBB7AB-AC7B-4F3D-A091-1238925E0448}
    string sComment = "备用"
  [41]
    dio dDio = {link=C3CF7374-59EF-4029-99B4-FC98E25808BB}
    string sComment = "备用"
  [42]
    dio dDio = {link=90C02E77-8235-444D-99EB-D816EF90AFE5}
    string sComment = "备用"
  [43]
    dio dDio = {link=E44556E2-741A-40A0-89B2-8E32677B3EB1}
    string sComment = "备用"
  [44]
    dio dDio = {link=D8AFCC23-6F61-4ADD-8DE3-3FE1547AD28D}
    string sComment = "备用"
  [45]
    dio dDio = {link=98BC2888-38BC-4A33-A762-BDEC3E36173F}
    string sComment = "备用"
  [46]
    dio dDio = {link=A24DA26D-2F10-46AE-809B-0B04336865AA}
    string sComment = "备用"
  [47]
    dio dDio = {link=04D21FA2-EBE1-4E66-8338-7CB17174A724}
    string sComment = "备用"
  [48]
    dio dDio = {link=E766472B-9569-4911-A858-6F7708718D01}
    string sComment = "备用"
  [49]
    dio dDio = {link=92C360C1-157E-40E1-9184-03D53ECDF3F7}
    string sComment = "备用"
  [50]
    dio dDio = {link=6E33B145-BAC8-48E7-A184-E5A9D90B515B}
    string sComment = "备用"
  [51]
    dio dDio = {link=D5FDB290-CB76-4852-8AF4-F9B6FA5D3E2D}
    string sComment = "备用"
  [52]
    dio dDio = {link=547C3630-B2EA-42F8-AB37-EEB4C81AA149}
    string sComment = "备用"
  [53]
    dio dDio = {link=A60C469C-4F75-4C30-9347-66365041DE79}
    string sComment = "备用"
  [54]
    dio dDio = {link=6E14BCEF-8B69-4038-B259-0EF712D2AB66}
    string sComment = "备用"
  [55]
    dio dDio = {link=B19F0E1B-CE25-49C3-9ED7-92404708DBC9}
    string sComment = "备用"
  [56]
    dio dDio = {link=AFC49D6D-7F53-41F5-8159-6058E9291542}
    string sComment = "备用"
  [57]
    dio dDio = {link=BB08126F-937C-4C50-9A1C-252CB13BB25C}
    string sComment = "备用"
  [58]
    dio dDio = {link=15BF4171-EFAA-47B7-BEF9-A698BE11011C}
    string sComment = "备用"
  [59]
    dio dDio = {link=9A261803-1F52-41D2-8355-1C79BF1BB94D}
    string sComment = "备用"
  [60]
    dio dDio = {link=18F63136-91BD-4FEE-8DA3-2AA9D2E8FFA8}
    string sComment = "备用"
  [61]
    dio dDio = {link=55E89D2C-C808-4026-99D2-85E324C475F9}
    string sComment = "备用"
  [62]
    dio dDio = {link=45535323-0512-46DB-8EB0-4BF3F55D73C7}
    string sComment = "备用"
  [63]
    dio dDio = {link=23943399-CEE5-49D9-BFD9-55B5920F548B}
    string sComment = "备用"
  [64]
    dio dDio = {link=364F41EB-6BA1-4700-BD0A-C2236839044E}
    string sComment = "备用"
  [65]
    dio dDio = {link=96EFCAAE-6B9A-4070-B9EC-2035BA94CCB3}
    string sComment = "备用"
  [66]
    dio dDio = {link=FD79DB68-803F-47E7-8305-8CFFFE519C88}
    string sComment = "备用"
  [67]
    dio dDio = {link=82CF98E3-5511-4523-9501-B4BBAD9DC96D}
    string sComment = "备用"
  [68]
    dio dDio = {link=43A446B7-3C25-4DD5-9597-27365DBE2539}
    string sComment = "备用"
  [69]
    dio dDio = {link=01367322-9745-4163-BFB8-DF881D521F4A}
    string sComment = "备用"
  [70]
    dio dDio = {link=1F635259-38C5-4AB2-B093-ADA4F82FD92B}
    string sComment = "备用"
  [71]
    dio dDio = {link=80065B3A-E7EF-4B6D-A30A-AC2F8A1FF9BD}
    string sComment = "备用"
  [72]
    dio dDio = {link=138692BF-FCCE-4B34-B0E8-8C4B22C67F12}
    string sComment = "备用"
  [73]
    dio dDio = {link=2F598E66-6704-43A6-A433-14D902C15D10}
    string sComment = "备用"
  [74]
    dio dDio = {link=3D7C9642-411B-40D3-B3B9-C83D24259AF4}
    string sComment = "备用"
  [75]
    dio dDio = {link=2E14C0AE-1F04-4256-8959-DEAD28BB69AE}
    string sComment = "备用"
  [76]
    dio dDio = {link=D90512A1-D0E1-41B2-8294-59D7C1ADD8E0}
    string sComment = "备用"
  [77]
    dio dDio = {link=F9EFA2A2-C655-4B55-8F3F-AAE77A6FD751}
    string sComment = "备用"
  [78]
    dio dDio = {link=8C43F822-1313-4C63-84D2-76D62B96A58F}
    string sComment = "备用"
  [79]
    dio dDio = {link=0BE51982-5E8E-4776-A637-0836608FA4D4}
    string sComment = "备用"
  [80]
    dio dDio = {link=5CC26A0C-A759-4F9D-9C90-7643106A4280}
    string sComment = "备用"
  [81]
    dio dDio = {link=6B2348DB-D0C3-44B1-96EA-09FBC0D6D1F3}
    string sComment = "备用"
  [82]
    dio dDio = {link=091DC27E-E2EB-463E-8E4B-08B48E663650}
    string sComment = "备用"
  [83]
    dio dDio = {link=EC5520D5-F711-48B3-AE90-97344DDBEE5C}
    string sComment = "备用"
  [84]
    dio dDio = {link=E02811C8-C36E-4E92-B28C-81A727813C5B}
    string sComment = "备用"
  [85]
    dio dDio = {link=39EB69C5-9612-415D-9A77-D013E3B8CFD4}
    string sComment = "备用"
  [86]
    dio dDio = {link=FD4FFC3C-593A-4304-8BB2-18534DB95237}
    string sComment = "备用"
  [87]
    dio dDio = {link=D2ECCFF1-C6D1-48A4-B3A9-F333711A9798}
    string sComment = "备用"
  [88]
    dio dDio = {link=13EA7043-3380-41E5-9177-AAC787C21C39}
    string sComment = "备用"
  [89]
    dio dDio = {link=5475660F-31B7-47C3-808C-FBAB066EFE6D}
    string sComment = "备用"
  [90]
    dio dDio = {link=93D7CC16-1244-4B9F-85C2-564B516A38A6}
    string sComment = "备用"
  [91]
    dio dDio = {link=A2A5B44E-CAC8-47F1-A810-875EED5095FB}
    string sComment = "备用"
  [92]
    dio dDio = {link=2F9951E4-3414-412E-A45B-55B5D632DA1B}
    string sComment = "备用"
  [93]
    dio dDio = {link=916866A1-8E9C-42B7-A695-7CB9D795E148}
    string sComment = "备用"
  [94]
    dio dDio = {link=CA3200CB-BA9D-4435-B593-6CDDBB86F10C}
    string sComment = "备用"
  [95]
    dio dDio = {link=49AC3AF5-F49B-42A1-90B2-5DB7D6C7E051}
    string sComment = "备用"
  [96]
    dio dDio = {link=64E7B72A-8AE1-43E7-9A21-FF4DABD03910}
    string sComment = "备用"
  [97]
    dio dDio = {link=7BA0757A-43B7-4994-86FC-1740DE8C159E}
    string sComment = "备用"
  [98]
    dio dDio = {link=5ACF5B88-9BD6-435A-8F3F-752FE88E7935}
    string sComment = "备用"
  [99]
    dio dDio = {link=70DFB9C6-9CA4-44C9-8464-A31BA0D039F5}
    string sComment = "备用"
  [100]
    dio dDio = {link=55D5D0F9-E23A-40DA-9955-6BCB63B37099}
    string sComment = "备用"
  [101]
    dio dDio = {link=1AB52030-AE2C-417B-9C38-1633EF57A0DB}
    string sComment = "备用"
  [102]
    dio dDio = {link=FFE2E20E-ABB5-4A36-BE3B-E714CB40E85A}
    string sComment = "备用"
  [103]
    dio dDio = {link=83BC89DD-B780-47A7-BBF0-017BDC2BA365}
    string sComment = "备用"
  [104]
    dio dDio = {link=10D6F5C6-79FE-4371-9CC9-A814346F77C1}
    string sComment = "备用"
  [105]
    dio dDio = {link=240957B0-B56A-4DFB-9281-23480961F3F1}
    string sComment = "备用"
  [106]
    dio dDio = {link=92C2EE73-BB65-4A97-8029-77FB60FFC23C}
    string sComment = "备用"
  [107]
    dio dDio = {link=62C2F98E-E7EB-49ED-971A-83A5444F6152}
    string sComment = "备用"
  [108]
    dio dDio = {link=58CC62E1-4595-401C-8E2F-3122D818CC74}
    string sComment = "备用"
  [109]
    dio dDio = {link=6D2EBC96-6FF5-40C1-83D6-CC8DD3D9FC3A}
    string sComment = "备用"
  [110]
    dio dDio = {link=AEC5DD07-0ABE-4FC2-A89A-ED52FEBBCAD7}
    string sComment = "备用"
  [111]
    dio dDio = {link=D289FF49-1CD8-4174-B7A5-8E375EB48B35}
    string sComment = "备用"
  [112]
    dio dDio = {link=4D3459D2-B2AE-4602-8654-6AD44AA154CE}
    string sComment = "备用"
  [113]
    dio dDio = {link=BE4318FA-0CA3-4B50-ACFD-D0BD90E002BB}
    string sComment = "备用"
  [114]
    dio dDio = {link=03734564-3942-45B2-807F-C861E4A00B4D}
    string sComment = "备用"
  [115]
    dio dDio = {link=18C4B14F-9C0F-4159-B56F-314AFF4BFABC}
    string sComment = "备用"
  [116]
    dio dDio = {link=A703F976-FEB8-4965-8F5A-CAD8585E54F7}
    string sComment = "备用"
  [117]
    dio dDio = {link=F3814F6C-1F81-45E4-8DE4-AB9F0C1AC9C1}
    string sComment = "备用"
  [118]
    dio dDio = {link=CD215C83-5C8C-4339-BF6C-DDE6EDBF5021}
    string sComment = "备用"
  [119]
    dio dDio = {link=295A35FF-B8CC-4A25-BC99-5CC4EFE79E3D}
    string sComment = "备用"
  [120]
    dio dDio = {link=7D822E1A-7C34-46E1-A06C-E10F3FD6B4DE}
    string sComment = "备用"
  [121]
